
// ===== library types =====

// folder: IO-Link Datatypes/3SU1 IDKey Switch

TYPE "LIOLink_3SU1_IDKeySwitch_typePII"
VERSION : 0.1
   STRUCT
      Status : Byte;
      IDKeyPlugged : Bool;
      AuthLvl_BIT0 : Bool;
      AuthLvl_BIT1 : Bool;
      AuthLvl_BIT2 : Bool;
      SwitchPos_BIT0 : Bool;
      SwitchPos_BIT1 : Bool;
      SwitchPos_BIT2 : Bool;
      Reserved : Bool;
   END_STRUCT;
END_TYPE

// folder: IO-Link ProzessData

TYPE "LIOLink_RF200_typePII"
TITLE = RFID_PII
VERSION : 0.1
   STRUCT
      UID : Array[0..7] of Byte;   // UID capturing / UID Erfassung
   END_STRUCT;
END_TYPE

TYPE "LIOLink_RF200_typePIQ"
TITLE = RFID_PIQ
VERSION : 0.1
   STRUCT
      AntennaOnOff : Byte;   // Antenna switch off with 16#10 (Bit 4 = TRUE) / Antenne ausschalten mit 16#10 (Bit 4 = TRUE)
      reserved : Array[0..6] of Byte;   // Reserved / Reserviert
   END_STRUCT;
END_TYPE

TYPE "LIOLink_3RR24_typePIQ"
TITLE = 3RR24_PIQ
VERSION : 0.1
   STRUCT
      StartOnDelayTime : Bool;   // Start On-Delay time / Starte Anlaufverzögerungszeit
      DQx1 : Bool;   // reserved / Reserviert
      DQx2 : Bool;   // reserved / Reserviert
      Reset : Bool;   // Reset
      DQx4 : Bool;   // reserved / Reserviert
      DQx5 : Bool;   // reserved / Reserviert
      DQx6 : Bool;   // reserved / Reserviert
      DQx7 : Bool;   // reserved / Reserviert
      DQx8 : Bool;   // reserved / Reserviert
      DQx9 : Bool;   // reserved / Reserviert
      DQx10 : Bool;   // reserved / Reserviert
      DQx11 : Bool;   // reserved / Reserviert
      DQx12 : Bool;   // reserved / Reserviert
      DQx13 : Bool;   // reserved / Reserviert
      DQx14 : Bool;   // reserved / Reserviert
      DQx15 : Bool;   // reserved / Reserviert
   END_STRUCT;
END_TYPE

TYPE "LIOLink_3RS1_typePIQ"
TITLE = 3RS14_PIQ
VERSION : 0.1
   STRUCT
      StartOnDelayTime : Bool;   // Start On-Delay time / Starte Anlaufverzögerungszeit
      DQx1 : Bool;   // reserved / Reserviert
      DQx2 : Bool;   // reserved / Reserviert
      Reset : Bool;   // Reset
      DQx4 : Bool;   // reserved / Reserviert
      DQx5 : Bool;   // reserved / Reserviert
      DQx6 : Bool;   // reserved / Reserviert
      DQx7 : Bool;   // reserved / Reserviert
      DQx8 : Bool;   // reserved / Reserviert
      DQx9 : Bool;   // reserved / Reserviert
      DQx10 : Bool;   // reserved / Reserviert
      DQx11 : Bool;   // reserved / Reserviert
      DQx12 : Bool;   // reserved / Reserviert
      DQx13 : Bool;   // reserved / Reserviert
      DQx14 : Bool;   // reserved / Reserviert
      DQx15 : Bool;   // reserved / Reserviert
   END_STRUCT;
END_TYPE

TYPE "LIOLink_3UG48_typePIQ"
TITLE = 3UG48_PIQ
VERSION : 0.1
   STRUCT
      StartTime : Bool;   // Start stabilization or On-Delay time / Starte Stabilisierungs- oder Anlaufverzögerungszeit
      DQx1 : Bool;   // reserved / Reserviert
      DQx2 : Bool;   // reserved / Reserviert
      Reset : Bool;   // Reset
      DQx4 : Bool;   // reserved / Reserviert
      DQx5 : Bool;   // reserved / Reserviert
      DQx6 : Bool;   // reserved / Reserviert
      DQx7 : Bool;   // reserved / Reserviert
      DQx8 : Bool;   // reserved / Reserviert
      DQx9 : Bool;   // reserved / Reserviert
      DQx10 : Bool;   // reserved / Reserviert
      DQx11 : Bool;   // reserved / Reserviert
      DQx12 : Bool;   // reserved / Reserviert
      DQx13 : Bool;   // reserved / Reserviert
      DQx14 : Bool;   // reserved / Reserviert
      DQx15 : Bool;   // reserved / Reserviert
   END_STRUCT;
END_TYPE

TYPE "LIOLink_3RR24_typePII"
TITLE = 3RR24_PII
VERSION : 0.1
// Das Prozessabbild der Eingänge enthält die wichtigsten Statusinformationen der
// Stromüberwachungsrelais 3RR24.
   STRUCT
      Rdy : Bool;   // Ready / Betriebsbereit
      DIx1 : Bool;   // reserved / Reserviert
      GroupError : Bool;   // Group error / Sammelfehler
      GroupWarning : Bool;   // Group warning / Sammelwarnung
      K1 : Bool;   // Status output relay K1 / Status Ausgangrelais K1
      DIx5 : Bool;   // reserved / Reserviert
      DIx6 : Bool;   // reserved / Reserviert
      DIx7 : Bool;   // reserved / Reserviert
      AnalogValueCoding : Byte;   // Analog value coding (only Bit 0..5) / Analogwertcodierung (nur Bit 0..5)
      AnalogValue : Int;   // Analog value / Analogwert
   END_STRUCT;
END_TYPE

TYPE "LIOLink_3UG48_typePII"
TITLE = 3UG48_PII / 3RR24_PII
VERSION : 0.1
// Das Prozessabbild der Eingänge enthält die wichtigsten Statusinformationen der
// Stromüberwachungsrelais 3RR24.
   STRUCT
      Rdy : Bool;   // Ready / Betriebsbereit
      DIx1 : Bool;   // reserved / Reserviert
      GroupError : Bool;   // Group error / Sammelfehler
      GroupWarning : Bool;   // General or group warning / Sammelwarnung
      K1 : Bool;   // Status output relay K1 / Status Ausgangrelais K1
      DIx5 : Bool;   // reserved / Reserviert
      DIx6 : Bool;   // reserved / Reserviert
      DIx7 : Bool;   // reserved / Reserviert
      AnalogValueCoding : Byte;   // Analog value coding (only Bit 0..5) / Analogwertcodierung (nur Bit 0..5)
      AnalogValue : Int;   // Analog value / Analogwert
   END_STRUCT;
END_TYPE

TYPE "LIOLink_3RA_typePII"
TITLE = 3RAxy_PII
VERSION : 0.1
// Data Type of the process input image contains the important status information of all compact starters. / Datentyp für das Prozessabbild der Eingänge enthält die wichtigen Statusinformationen aller Kompaktabzweige.
   STRUCT
      St1Rdy : Bool;   // Starter 1 ready (automatic) / Starter 1 Bereit (Automatik)
      St1MotorOn : Bool;   // Starter 1 Motor on / Starter 1 Motor ein
      St1Fault : Bool;   // Starter 1 group fault / Starter 1 Sammelfehler
      St1Warn : Bool;   // Starter 1 group warning / Starter 1 Sammelwarnung
      St2Rdy : Bool;   // Starter 2 ready (automatic) / Starter 2 Bereit (Automatik)
      St2MotorOn : Bool;   // Starter 2 Motor on / Starter 2 Motor ein
      St2Fault : Bool;   // Starter 2 group fault / Starter 2 Sammelfehler
      St2Warn : Bool;   // Starter 2 group warning / Starter 2 Sammelwarnung
      St3Rdy : Bool;   // Starter 3 ready (automatic) / Starter 3 Bereit (Automatik)
      St3MotorOn : Bool;   // Starter 3 Motor on / Starter 3 Motor ein
      St3Fault : Bool;   // Starter 3 group fault / Starter 3 Sammelfehler
      St3Warn : Bool;   // Starter 3 group warning / Starter 3 Sammelwarnung
      St4Rdy : Bool;   // Starter 4 ready (automatic) / Starter 4 Bereit (Automatik)
      St4MotorOn : Bool;   // Starter 4 Motor on / Starter 4 Motor ein
      St4Fault : Bool;   // Starter 4 group fault / Starter 4 Sammelfehler
      St4Warn : Bool;   // Starter 4 group warning / Starter 4 Sammelwarnung
   END_STRUCT;
END_TYPE

TYPE "LIOLink_3RA_typePIQ"
TITLE = 3RAxy_PIQ
VERSION : 0.1
// The process output image contains the control commands for all compact starters. / Datentyp für das Prozessabbild der Ausgänge enthält die Steuerbefehle für alle Kompaktabzweige.
   STRUCT
      St1Dir1 : Bool;   // Starter 1 Motor direction of rotation 1 / Starter 1 Motor Drehrichtung 1
      St1Dir2 : Bool;   // Starter 1 Motor direction of rotation 2 / Starter 1 Motor Drehrichtung 2
      St1Res : Bool;   // Starter 1 Reserved / Starter 1 reserviert
      St1TripReset : Bool;   // Starter 1 Trip reset / Starter 1 Trip-Reset
      St2Dir1 : Bool;   // Starter 2 Motor direction of rotation 1 / Starter 2 Motor Drehrichtung 1
      St2Dir2 : Bool;   // Starter 2 Motor direction of rotation 2 / Starter 2 Motor Drehrichtung 2
      St2Res : Bool;   // Starter 2 Reserved / Starter 2 reserviert
      St2TripReset : Bool;   // Starter 2 Trip reset / Starter 2 Trip-Reset
      St3Dir1 : Bool;   // Starter 3 Motor direction of rotation 1 / Starter 3 Motor Drehrichtung 1
      St3Dir2 : Bool;   // Starter 3 Motor direction of rotation 2 / Starter 3 Motor Drehrichtung 2
      St3Res : Bool;   // Starter 3 Reserved / Starter 3 reserviert
      St3TripReset : Bool;   // Starter 3 Trip reset / Starter 3 Trip-Reset
      St4Dir1 : Bool;   // Starter 4 Motor direction of rotation 1 / Starter 4 Motor Drehrichtung 1
      St4Dir2 : Bool;   // Starter 4 Motor direction of rotation 2 / Starter 4 Motor Drehrichtung 2
      St4Res : Bool;   // Starter 4 Reserved / Starter 4 reserviert
      St4TripReset : Bool;   // Starter 4 Trip reset / Starter 4 Trip-Reset
   END_STRUCT;
END_TYPE

TYPE "LIOLink_3RB24_typePII"
TITLE = 3RB24_PII
VERSION : 0.1
// Data Type of the process input image contains the most important status information of the solid-state overload relay for IO‑Link.
// Datentyp für das Prozessabbild der Eingänge enthält die wichtigsten Statusinformationen des
// elektronischen Überlastrelais für IO-Link.
   STRUCT
      Rdy : Bool;   // Ready (automatic) / Bereit (Automatik)
      MotorOn : Bool;   // Motor on / Motor ein
      GroupFault : Bool;   // Group fault / Sammelfehler
      GroupWarning : Bool;   // Group warning / Sammelwarnung
      DIx4 : Bool;   // reserved / reserviert
      DIx5 : Bool;   // reserved / reserviert
      DIx6 : Bool;   // reserved / reserviert
      DIx7 : Bool;   // reserved / reserviert
      CurrentRatio : Byte;   // Bit 0..5: Motor current ratio (%), Bit 6: Manual mode / Bit 0..5: Motorstromverhältnis, Bit 6: Handbetrieb
   END_STRUCT;
END_TYPE

TYPE "LIOLink_3RB24_typePIQ"
TITLE = 3RB24_PIQ
VERSION : 0.1
// The process output image contains the control commands for the solid-state overload relay for IO‑Link.
// Datentyp für das Prozessabbild der Ausgänge enthält die Steuerbefehle für das elektronische
// Überlastrelais für IO-Link
   STRUCT
      Direction1 : Bool;   // Motor direction of rotation 1 / Motor Drehrichtung 1
      Direction2 : Bool;   // Motor direction of rotation 2 / Motor Drehrichtung 2
      DQx2 : Bool;   // Reserved / reserviert
      TripReset : Bool;   // Trip reset / Trip-Reset
      DQx4 : Bool;   // Reserved / reserviert
      DQx5 : Bool;   // Reserved / reserviert
      DQx6 : Bool;   // Reserved / reserviert
      DQx7 : Bool;   // Reserved / reserviert
      DQx8 : Bool;   // Reserved / reserviert
      DQx9 : Bool;   // Reserved / reserviert
      DQx10 : Bool;   // Reserved / reserviert
      DQx11 : Bool;   // Reserved / reserviert
      DQx12 : Bool;   // Reserved / reserviert
      DQx13 : Bool;   // Reserved / reserviert
      DQx14 : Bool;   // Reserved / reserviert
      DQx15 : Bool;   // Reserved / reserviert
   END_STRUCT;
END_TYPE

TYPE "LIOLink_3RS1_typePII"
TITLE = 3RS14_PII
VERSION : 0.1
   STRUCT
      Rdy : Bool;   // Ready / Betriebsbereit
      DIx1 : Bool;   // reserved / Reserviert
      GroupError : Bool;   // Group error / Sammelfehler
      GroupWarning : Bool;   // General or group warning / Sammelwarnung
      K1 : Bool;   // Status output relay K1 / Status Ausgangrelais K1
      K2 : Bool;   // Status output relay K2 / Status Ausgangrelais K2
      K3 : Bool;   // Status output relay K3 / Status Ausgangrelais K3
      DIx7 : Bool;   // reserved / Reserviert
      AnalogValueCoding : Byte;   // Analog value coding (only Bit 0..4) / Analogwertcodierung (nur Bit 0..4)
      AnalogValue : Int;   // Analog value / Analogwert
   END_STRUCT;
END_TYPE

// folder: LIOLink

TYPE "LIOLink_typeDiagnostics"
   STRUCT
      status : Word;   // Status of the Block or error identification when error occurred
      subfunctionStatus : DWord;   // Status or return value of called FB's, FCs and system blocks
      stateNumber : DInt;   // State in the state machine of the block where the error occurred
   END_STRUCT;
END_TYPE

// folder: LIOLink/Common

TYPE "LIOLink_typePortEventQualifier"
TITLE = LIOLink_typePortEventQualifier
// EventQualifier: Instance, Source, Type, Mode
   STRUCT
      instance : Byte;   // 0: Unknown / 1-3: Reserved / 4: Application / 5-7: Reserved
      source : Bool;   // (default) FALSE: Device (remote) / TRUE: Master/Port
      "type" : Byte;   // 0: Reserved / 1: Notification / 2: Warning / 3: Error
      mode : Byte;   // 0: Reserved / 1: Event single shot / 2: Event disappears / 3: Event appears
   END_STRUCT;
END_TYPE

TYPE "LIOLink_typePortEventCodes"
TITLE = LIOLink_PortEventCodes
// UDT for Event Information: eventCode, eventQualifier
   STRUCT
      eventCode : Word;   // IO-Link EventCode
      eventQualifier : "LIOLink_typePortEventQualifier";   // IO-Link EventQualifier
   END_STRUCT;
END_TYPE

TYPE "LIOLink_typePortEvents"
TITLE = LIOLink_PortEvents
// Events of a port
   STRUCT
      event : Array[0..4] of "LIOLink_typePortEventCodes";   // Events of a port
   END_STRUCT;
END_TYPE

TYPE "LIOLink_typeEvents"
TITLE = LIOLink_Events
// Events of each port of a IO-Link-Master
   STRUCT
      port : Array[1..8] of "LIOLink_typePortEvents";   // Ports of IO-Link-Master
   END_STRUCT;
END_TYPE

// folder: LIOLink/Common/Device-specific data types/SIMATIC RF200

TYPE "LIOLink_RF200_typeParameters"
TITLE = LIOLink_RF200_typeParameters
// Contains all parameters of a RF200
   STRUCT
      eventMessage : Byte;   // 16#02: Event indication enabled (default), 16#04: No Message
      operatingMode : Byte;   // 16#04: Scan UID (default), 16#08 Scan user data
      readyDelay : Byte;   // 16#02 Turn off (default), 16#04: Turn on additional backup mechanism for
      dataHoldingTime : Byte;   // Minimum time during which the process input data is not changed by the device
      rfParameters : Byte;   // Setting the RF parameters, 16#02 ISO default, 16#04: special settings
      modulation : Byte;   // Setting for the modulation strength 16#00 (0%) ... 16#64 (100%) - default 16#16 (22%)
      subcarrier : Byte;   // Subcarrier, 16#02: Single (default), 16#04: double
      dataTransfer : Byte;   // Data transmission speed, 16#02: low, 16#04: high (default)
   END_STRUCT;
END_TYPE

TYPE "LIOLink_RF200_typeEventHistory"
TITLE = LIOLink_RF200_typeEventHistory
VERSION : 0.1
// Contains last 5 events of a RF200
   STRUCT
      lastEvent : DWord;   // Last event
      secondLastEvent : DWord;   // Second last event
      thirdLastEvent : DWord;   // Third last event
      fourthLastEvent : DWord;   // Fourth last event
      fifthLastEvent : DWord;   // Fifth last event
   END_STRUCT;
END_TYPE

TYPE "LIOLink_RF200_typeReaderStatus"
TITLE = LIOLink_RF200_typeReaderStatus
VERSION : 0.1
// Contrains all information about the status of the reader
   STRUCT
      timeSinceStartup : DWord;   // Operating time in seconds
      tagsInTheField : Byte;   // current number of transponders in the field
      antennaStatus : Byte;   // antenna turned on/off
      tagChanges : DWord;   // number of transponder changes
      lineDriverRev : Byte;   // version of the IO-Link line driver
      errorCounterPassive : Byte;   // Air interface: Counter for errors in idle state
      abortCounter : Byte;   // Air interface: Communication aborted
      codeErrorCounter : Byte;   // Air interface: Communication disruption
      signatureErrorCounter : Byte;   // Air interface: Protocol error, signature error counter, is reset when read out
      crcErrorCounter : Byte;   // Air interface: Communication disruption
      currentCommandStatus : Byte;   // Command status of the last command, is reset when read out
      errorCount : Byte;   // HOST interface: Communication disruption
   END_STRUCT;
END_TYPE

TYPE "LIOLink_RF200_typeUIDHistory"
TITLE = LIOLink_RF200_typeUIDHistory
VERSION : 0.1
// Contains UID history
   STRUCT
      lastUID1 : DWord;   // Last UID
      lastUID2 : DWord;   // Last UID
      secondLastUID1 : DWord;   // Second last UID
      secondLastUID2 : DWord;   // Second last UID
      thirdLastUID1 : DWord;   // Third last UID
      thirdLastUID2 : DWord;   // Third last UID
      fourthLastUID1 : DWord;   // Fourth last UID
      fourthLastUID2 : DWord;   // Fourth last UID
      fifthLastUID1 : DWord;   // Fifth last UID
      fifthLastUID2 : DWord;   // Fifth last UID
   END_STRUCT;
END_TYPE

TYPE "LIOLink_RF200_typeTagStatus"
TITLE = LIOLink_RF200_typeTagStatus
VERSION : 0.1
// Contains all the information about the status of the tag
   STRUCT
      uid : Array[0..7] of Byte;   // Unique identifier of the transponder
      tagName : Byte;   // Transponder Name
      chipVersion : Byte;   // Version of the Chip
      memSize : Word;   // Memory size in Bytes
      lockStatus : Byte;   // Disable blocks on the chip
      memBlockSize : Byte;   // Size of memory blocks of the chip
      numBlocks : Byte;   // Number of memory blocks of the chip
   END_STRUCT;
END_TYPE

TYPE "LIOLink_RF200_typeAll"
TITLE = LIOLink_RF200_typeAll
VERSION : 0.1
// Contains all information about RF200
   STRUCT
      directParameterPage : "LIOLink_typeParameterPage0";   // ID0: Parameter page 0
      systemCommand : Byte;   // ID2: System command
      deviceAccessLocks : Word;   // ID12: Device access locks
      vendorName : String[12];   // ID16: Vendor name
      vendorText : String[12];   // ID17: Vendor text
      productName : String[24];   // ID18: Product name
      productID : String[16];   // ID19: Product ID
      productText : String[64];   // ID20: Product Text
      serialNumber : String[12];   // ID21: Serial Number
      hwRevision : String[12];   // ID22: Hardware revision
      fwRevision : String[12];   // ID23: Firmware revision
      appSpecificName : String[32];   // ID24: Application specific name
      errorCount : Word;   // ID32: Number of errors that have occured (not warnings)
      deviceStatus : Byte;   // ID36: Device status
      deviceStatusDetailed : Byte;   // ID37: Detailed device status
      processImageIn : Array[0..7] of Byte;   // ID40: Read out last process image of the inputs
      processImageOut : Array[0..7] of Byte;   // ID41: Read out last process image of the outputs
      parameters : "LIOLink_RF200_typeParameters";   // ID64: Read/Write Reader Parameters
      eventHistory : "LIOLink_RF200_typeEventHistory";   // ID74: Number of events
      readerStatus : "LIOLink_RF200_typeReaderStatus";   // ID90: Reader status
      tagStatus : "LIOLink_RF200_typeTagStatus";   // ID91: Tag status
      uidHistory : "LIOLink_RF200_typeUIDHistory";   // ID92: History of UID
   END_STRUCT;
END_TYPE

// folder: LIOLink/Common/Device-specific data types/SIRIUS/3RA

TYPE "LIOLink_3RA_typeDiagStarterShort"
TITLE = LIOLink_3RA_typeDiagStarterShort
// Contains diagnose of starter of type "short"
   STRUCT
      starterItemNumber : Byte;   // Starter Item number (1 to 4)
      starterAvailable : Byte;   // Starter Available: 16#00 not available; 16#02: available
      reserved1 : Array[2..5] of Byte;   // Reserved
      contactBlockDefective : Bool;   // Contact block defective
      contactSupplyVoltageMissing : Bool;   // Contact block supply voltage missing
      reserved2 : Bool;   // Reserved
      trippMotorOverload : Bool;   // Motor overload tripping
      trippCircuitBreaker : Bool;   // Circuit breaker tripped
      switchOffendPosRight : Bool;   // Switch off - end position right
      switchOffendPosLeft : Bool;   // Switch off - end position left
      processImageError : Bool;   // Process image error
      manualOperationLocal : Bool;   // Manual operation local
      manualOperationConAborted : Bool;   // Manual operation connection aborted
      ContactCoolingTimeActive : Bool;   // Contact block cooling time active
      remainingLifeTime0 : Bool;   // Remaining life time (RLT 0%)
      reserved3 : Bool;   // Reserved
      reserved4 : Bool;   // Reserved
      reserved5 : Bool;   // Reserved
      reserved6 : Bool;   // Reserved
   END_STRUCT;
END_TYPE

TYPE "LIOLink_3RA_typeDiagStarterLong"
TITLE = LIOLink_3RA_typeDiagStarterLong
// Contains diagnose of starter of type "long"
   STRUCT
      reserved1 : Byte;   // Reserved
      starterItemNumber : Byte;   // Starter Item number (1 to 4)
      starterAvailable : Byte;   // Starter Available: 16#00 not available; 16#02: available
      reserved2 : Array[3..6] of Byte;   // Reserved
      contactBlockDefective : Bool;   // Contact block defective
      contactSupplyVoltageMissing : Bool;   // Contact block supply voltage missing
      reserved3 : Bool;   // Reserved
      trippMotorOverload : Bool;   // Motor overload tripping
      trippCircuitBreaker : Bool;   // Circuit breaker tripped
      switchOffendPosRight : Bool;   // Switch off - end position right
      switchOffendPosLeft : Bool;   // Switch off - end position left
      processImageError : Bool;   // Process image error
      manualOperationLocal : Bool;   // Manual operation local
      manualOperationConAborted : Bool;   // Manual operation connection aborted
      ContactCoolingTimeActive : Bool;   // Contact block cooling time active
      remainingLifeTime0 : Bool;   // Remaining life time (RLT 0%)
      reserved4 : Bool;   // Reserved
      reserved5 : Bool;   // Reserved
      reserved6 : Bool;   // Reserved
      reserved7 : Bool;   // Reserved
      reserved8 : Byte;   // Reserved
   END_STRUCT;
END_TYPE

TYPE "LIOLink_3RA_typeConfigStarterShort"
TITLE = LIOLink_3RA_typeConfigStarterShort
// Contains configurations for starter with type "short"
   STRUCT
      starterItemNumber : Byte;   // Starter (item number)
      reserved1 : Byte := 16#60;   // Fixed Value
      starterDiag : Byte;   // Starter Diag: 16#00: not available; 16#02: available but defect; 16#03: available and OK
      starterType : Byte;   // Type of starter
      starterVersion1 : Byte;   // Starter Version part 1
      starterVersion2 : Byte;   // Starter Version part 2
   END_STRUCT;
END_TYPE

TYPE "LIOLink_3RA_typeConfigStarterLong"
TITLE = LIOLink_3RA_typeConfigStarterLong
// Contains configurations for starter with type "long"
   STRUCT
      reserved : Byte := 16#07;   // Fixed Value
      starterItemNumber : Byte;   // Starter (item number)
      reserved1 : Byte := 16#60;   // Fixed Value
      starterDiag : Byte;   // Starter Diag: 16#00: not available; 16#02: available but defect; 16#03: available and OK
      starterType : Byte;   // Type of starter
      starterVersion1 : Byte;   // Starter Version part 1
      starterVersion2 : Byte;   // Starter Version part 2
      reserved2 : Byte := 16#07;   // Fixed Value
   END_STRUCT;
END_TYPE

TYPE "LIOLink_3RA_typeDiag"
TITLE = LIOLink_3RA_typeDiag
VERSION : 0.1
// Data set (index) 90 - group diagnostics: Starter group
   STRUCT
      reserved : Array[0..3] of Byte;   // Reserved - Dataset Index 90 - Length 53 / read length 52
      numberOfStarters : Byte;   // Number of starters (compact starters and operator panel)
      configurationCompare : Byte;   // Preset <> actual configuration 16#00: equal 16#01: different
      reserved1 : Word;   // Reserved
      starter1 : "LIOLink_3RA_typeDiagStarterLong";   // Starter 1 - module and specific diagnostics
      starter2 : "LIOLink_3RA_typeDiagStarterShort";   // Starter 2 - module and specific diagnostics
      starter3 : "LIOLink_3RA_typeDiagStarterLong";   // Starter 3 - module and specific diagnostics
      starter4 : "LIOLink_3RA_typeDiagStarterShort";   // Starter 4 - module and specific diagnostics
      reserved3 : Byte;   // Reserved
      operatorItemNumber : Byte;   // Operator panel (item number)
      operatorAvailable : Byte;   // Operator panel available: 16#00 not available; 16#02: available
      reserved4 : Byte;   // Reserved
      reserved5 : Array[48..51] of Byte;   // Reserved
   END_STRUCT;
END_TYPE

TYPE "LIOLink_3RA_typeConfig"
TITLE = LIOLink_3RA_typeConfig / IO-Link Parameter mit dem Baustein "FB IO_CALL" auslesen!
VERSION : 0.1
// Contains all the possible configurations of 3RA
   STRUCT
      reserved : Array[0..7] of Byte;   // Reserved
      starter1 : "LIOLink_3RA_typeConfigStarterLong";   // Config Data of Starter 1
      starter2 : "LIOLink_3RA_typeConfigStarterShort";   // Config Data of Starter 2
      starter3 : "LIOLink_3RA_typeConfigStarterLong";   // Config Data of Starter 3
      starter4 : "LIOLink_3RA_typeConfigStarterShort";   // Config Data of Starter 4
      reserved1 : Byte := 16#07;   // Reserved
      operatorItemNumber : Byte;   // Operator panel (item number)
      reserved2 : Byte := 16#60;   // Reserved
      operatorAvailable : Byte;   // Operator panel available: 16#00 not available; 16#02: available
      reserved3 : Byte := 16#D2;   // Reserved
      reserved4 : Byte;   // Reserved
   END_STRUCT;
   // reserved[0] := 16#0021;
   // reserved[1] := 16#0000;
   // reserved[2] := 16#0000;
   // reserved[3] := 16#0000;
   // reserved[4] := 16#0005;
END_TYPE

TYPE "LIOLink_3RA_typeAll"
TITLE = LIOLink_3RA_typeAll
VERSION : 0.1
// Contains all the information about 3RA
   STRUCT
      parameterPage0 : "LIOLink_typeParameterPage0";   // ID0: Parameter page 0
      parameterPage1 : "LIOLink_3RA_typeParameterPage1";   // ID1: Parameter page 1
      vendorName : String[10];   // ID16: Vendor name
      vendorText : String[58];   // ID17: Vendor text
      productName : String[30];   // ID18: Product name
      productID : String[8];   // ID19: Product ID
      productText : String[2];   // ID20: Product text
      serialNumber : String[8];   // ID21: Serial number
      hwRevision : String[4];   // ID22: Hardware revision
      fwRevision : String[4];   // ID23: Firmware revision
      appSpecificName : String[32];   // ID24: Application specific name
      diagnostics : "LIOLink_3RA_typeDiag";   // ID90: Group diagnostics
      actualConfig : "LIOLink_3RA_typeConfig";   // ID105: Actual configuration
      targetConfig : "LIOLink_3RA_typeConfig";   // ID130: Target configuration
   END_STRUCT;
   // actualConfig.reserved[0] := 16#0021;
   // actualConfig.reserved[1] := 16#0000;
   // actualConfig.reserved[2] := 16#0000;
   // actualConfig.reserved[3] := 16#0000;
   // actualConfig.reserved[4] := 16#0005;
   // targetConfig.reserved[0] := 16#0021;
   // targetConfig.reserved[1] := 16#0000;
   // targetConfig.reserved[2] := 16#0000;
   // targetConfig.reserved[3] := 16#0000;
   // targetConfig.reserved[4] := 16#0005;
END_TYPE

TYPE "LIOLink_3RA_typeParameterPage1"
TITLE = LIOLink_3RA_typeParameterPage1 / IO-Link Parameter mit dem Baustein "FB IO_CALL" auslesen!
AUTHOR : SIE_RS
FAMILY : 3RA
NAME : IO-Link
VERSION : 1.0
// Contains Parameter Page 1 of 3RA
   STRUCT
      productFamiliy : Byte;   // Produktfamily SIRIUS (0x60) - A-9 Dataset Index 1 Page 75
      starter1Compare : Bool;   // Starter 1 - 0: Target/actual comparison: Yes, 1: Target/actual comparison: No,
      starter1Available : Bool;   // Starter 1 - 0: Starter available: No, 1: Starter available: Yes,
      starter2Compare : Bool;   // Starter 2 - 0: Target/actual comparison: Yes, 1: Target/actual comparison: No,
      starter2Available : Bool;   // Starter 2 - 0: Starter available: No, 1: Starter available: Yes,
      starter3Compare : Bool;   // Starter 3 - 0: Target/actual comparison: Yes, 1: Target/actual comparison: No,
      starter3Available : Bool;   // Starter 3 - 0: Starter available: No, 1: Starter available: Yes,
      starter4Compare : Bool;   // Starter 4 - 0: Target/actual comparison: Yes, 1: Target/actual comparison: No,
      starter4Available : Bool;   // Starter 4 - 0: Starter available: No, 1: Starter available: Yes,
      operatorPanelCompare : Bool;   // Operator panel - 0:Target/actual comparison: Yes, 1:Target/actual comparison:No
      operatorPanelAvailable : Bool;   // Operator panel - 0: Starter available: No, 1: Starter available: Yes,
      reserved1 : Bool;   // Reserved
      reserved2 : Bool;   // Reserved
      profileVersion1 : Bool;   // Profile version
      profileVersion2 : Bool;   // Profile version
      profileVersion3 : Bool;   // Profile version
      profileVersion4 : Bool;   // Profile version
      starter1Type : Byte;   // Starter 1 - Type of starter
      starter1Version : Byte;   // Starter 1 - Starter version
      starter2Type : Byte;   // Starter 2 - Type of starter
      starter2Version : Byte;   // Starter 2 - Starter version
      starter3Type : Byte;   // Starter 3 - Type of starter
      starter3Version : Byte;   // Starter 3 - Starter version
      starter4Type : Byte;   // Starter 4 - Type of starter
      starter4Version : Byte;   // Starter 4 - Starter version
      operatorPanel : Byte;   // 210: Operator panel
      reserved3 : Byte;   // Reserved
      reserved4 : Byte;   // Reserved
      reserved5 : Byte;   // Reserved
      reserved6 : Byte;   // Reserved
   END_STRUCT;
END_TYPE

// folder: LIOLink/Common/Device-specific data types/SIRIUS/3RB24

TYPE "LIOLink_3RB24_typeMeasure"
TITLE = LIOLink_3RB24_typeMeasure
VERSION : 0.1
// Data set (index) 94 (measured values) - solid-state overload relay for IO‑Link
   STRUCT
      phaseCurrentL1Rel : Byte;   // Phase current I (L1 rms in 3,125% steps) - A-4 Dataset Index 94 Page 112
      phaseCurrentL2Rel : Byte;   // Phase current I (L2 rms in 3,125 % steps)
      phaseCurrentL3Rel : Byte;   // Phase current I (L3 rms in 3,125 % steps)
      reserved : Byte;   // Reserved
      reserved1 : Array[4..27] of Byte;   // Reserved
      phaseCurrentL1Abs : DWord;   // Phase current I (L1 rms in 0,01-A steps)
      phaseCurrentL2Abs : DWord;   // Phase current I (L2 rms in 0,01-A steps)
      phaseCurrentL3Abs : DWord;   // Phase current I (L3 rms in 0,01-A steps)
   END_STRUCT;
END_TYPE

TYPE "LIOLink_3RB24_typeTechFunctions"
TITLE = TechnologyFunctions_3RB24
VERSION : 0.1
// Data set (index) 131 (technology functions) - solid-state overload relay for IO‑Link
   STRUCT
      reserved : Array[0..7] of Byte;   // Reserved
      groundFaultDetection : Byte;   // Ground fault detection - 16#00: Disable; 16#20: Enable - Bit 5 in Byte
      reserved8 : Word;   // Reserved
      coldStart : Byte;   // Cold Start - 16#00: Disable; 16#08: Enable - Bit 3 in Byte
      ratedOpCurrent : DWord;   // Rated operational current (in 0.01 A steps)
      reserved16 : Word;   // Reserved
      responseToOverloadMotor : Byte;   // Response to overload - thermal motor model - 16#00: Tripping without restart (MAN); 16#01: Tripping with restart (AUTO)
      tripClass : Byte;   // Trip class - 16#03: CLASS 5; 16#00: CLASS 10; 16#01: CLASS 20; 16#02: CLASS 30
      reserved17 : DWord;   // Reserved
      responseToOverloadThermistor : Bool;   // Response to overload - Thermistor - false: Tripping without restart (MAN); true: Tripping with restart (AUTO)
      reserved18 : Bool;   // Reserved
      reserved19 : Bool;   // Reserved
      reserved20 : Bool;   // Reserved
      reserved21 : Bool;   // Reserved
      reserved22 : Bool;   // Reserved
      reserved23 : Bool;   // Reserved
      monitorThermistor : Bool;   // Thermistor - monitoring - false: No; true: Yes
   END_STRUCT;
END_TYPE

TYPE "LIOLink_3RB24_typePresetConfig"
TITLE = TargetConfiguration_3RB24
VERSION : 0.1
// Data set (index) 130 (target configuration) - operator panel
   STRUCT
      reserverd : Array[0..17] of Byte;   // Reserved
      reserved1 : Bool;   // Reserved
      reserved2 : Bool;   // Reserved
      reserved3 : Bool;   // Reserved
      reserved4 : Bool;   // Reserved
      reserved5 : Bool;   // Reserved
      reserved6 : Bool;   // Reserved
      operationAtTarget : Bool;   // Operation at Preset <> Actual Configuration
      operationPanelAvailable : Bool;   // Operator panel available
      reserved7 : Byte;   // Reserved
      reserved8 : Byte;   // Reserved
      reserved9 : Byte;   // Reserved
   END_STRUCT;
END_TYPE

TYPE "LIOLink_3RB24_typeDiag"
TITLE = LIOLink_3RB24_typeDiag
VERSION : 0.1
// Data set (index) 94 (measured values) - solid-state overload relay for IO‑Link
   STRUCT
      ready : Bool;   // Ready
      directionClockwise : Bool;   // Motor direction of rotation 1 (clockwise)
      directionCounterClockwise : Bool;   // Motor direction of rotation 2 (counter-clockwise)
      reserved : Bool;   // Reserved
      switchingElementDefect : Bool;   // Switching element defective
      reserved1 : Bool;   // Reserved
      groupError : Bool;   // GroupError
      generalWarning : Bool;   // General warning
      reserved2 : Byte;   // Reserved
      thermistorOverload : Bool;   // Thermistor overload
      thermistorWireBreak : Bool;   // Thermistor wire break
      thermistorShortCircuit : Bool;   // Thermistor short-circuit
      thermistorMotorOverload : Bool;   // Thermal motor model overload
      overloadTripping : Bool;   // Overload tripping
      reserved3 : Bool;   // Reserved
      reserved4 : Bool;   // Reserved
      reserved5 : Bool;   // Reserved
      reserved6 : Byte;   // Reserved
      reserved7 : Bool;   // Reserved
      reserved8 : Bool;   // Reserved
      reserved9 : Bool;   // Reserved
      reserved10 : Bool;   // Reserved
      reserved11 : Bool;   // Reserved
      resCurrenctDetected : Bool;   // Residual current detected
      resCurrentTripping : Bool;   // Residual current tripping
      reserved12 : Bool;   // Reserved
      reserved13 : Byte;   // Reserved
      groudFaultDetected : Bool;   // Ground fault detected
      GroundFaultTripping : Bool;   // Ground fault tripping
      reserved14 : Bool;   // Reserved
      reserved15 : Bool;   // Reserved
      reserved16 : Bool;   // Reserved
      reserved17 : Bool;   // Reserved
      reserved18 : Bool;   // Reserved
      supplyVoltageLow : Bool;   // Electronics supply voltage too low
      reserved19 : Bool;   // Reserved
      reserved20 : Bool;   // Reserved
      autoMode1 : Bool;   // Automatic mode
      autoMode2 : Bool;   // Automatic mode
      manualModeOP1 : Bool;   // Manual mode (operator panel)
      manualModeOP2 : Bool;   // Manual mode (operator panel)
      manualModeConAbort : Bool;   // Manual mode connection abort (operator panel)
      processImageError : Bool;   // Process image error
      reserved21 : Byte;   // Reserved
      selfTestActive1 : Bool;   // Self-test active
      selfTestActive2 : Bool;   // Self-test active
      selfTestError : Bool;   // Self-test error
      reserved22 : Bool;   // Reserved
      reserved23 : Bool;   // Reserved
      reserved24 : Bool;   // Reserved
      reserved25 : Bool;   // Reserved
      reserved26 : Bool;   // Reserved
      reserved27 : Word;   // Reserved
      reserved28 : Bool;   // Reserved
      reserved29 : Bool;   // Reserved
      impermissibleSetting : Bool;   // Impermissible Ie/CLASS setting
      presetActualCompare : Bool;   // Preset <> actual configuration
      thermistorProtectionDeactivated : Bool;   // Thermistor protection deactivated
      reserved30 : Bool;   // Reserved
      reserved31 : Bool;   // Reserved
      reserved32 : Bool;   // Reserved
      reserved33 : Byte;   // Reserved
      coldStartActive : Bool;   // Cold start active
      coldStartTripping : Bool;   // Cold start tripping
      reserved34 : Bool;   // Reserved
      reserved35 : Bool;   // Reserved
      reserved36 : Bool;   // Reserved
      reserved37 : Bool;   // Reserved
      reserved38 : Bool;   // Reserved
      reserved39 : Bool;   // Reserved
      reserved40 : Byte;   // Reserved
      reserved41 : Array[16..23] of Byte;   // Reserved
      reserved42 : Bool;   // Reserved
      reserved43 : Bool;   // Reserved
      reserved44 : Bool;   // Reserved
      motorHeatingExceeded : Bool;   // Prewarning limit: Motor heating exceeded
      reserved45 : Bool;   // Reserved
      reserved46 : Bool;   // Reserved
      reserved47 : Bool;   // Reserved
      reserved48 : Bool;   // Reserved
      reserved49 : Byte;   // Reserved - Extension to get even field
   END_STRUCT;
END_TYPE

TYPE "LIOLink_3RB24_typeAll"
TITLE = LIOLink_3RB24_typeAll
VERSION : 0.1
// Contains all the information about 3RB24
   STRUCT
      parameterPage0 : "LIOLink_typeParameterPage0";   // ID0: Parameter page 0
      vendorName : String[10];   // ID16: Vendor name
      vendorText : String[64];   // ID17: Vendor text
      productName : String[30];   // ID18: Product name
      productID : String[12];   // ID19: Product ID
      productText : String[2];   // ID20: Product text
      serialNumber : String[8];   // ID21: Serial number
      hwRevision : String[4];   // ID22: Hardware revision
      fwRevision : String[4];   // ID23: Firmware revision
      appSpecificName : String[32];   // ID24: Application specific name
      processInput : Word;   // ID40: Process data input
      processOutput : Byte;   // ID41: Process data output
      diagnostics : "LIOLink_3RB24_typeDiag";   // ID92: Diagnostics
      measuredValues : "LIOLink_3RB24_typeMeasure";   // ID94: Measurement values
      presetConfig : "LIOLink_3RB24_typePresetConfig";   // ID130: Preset configuration
      techFunctions : "LIOLink_3RB24_typeTechFunctions";   // ID131: Technology functions
   END_STRUCT;
END_TYPE

// folder: LIOLink/Common/Device-specific data types/SIRIUS/3RR24

TYPE "LIOLink_3RR24_typeDiag"
TITLE = LIOLink_3RR24_typeDiag
VERSION : 0.1
// Data set (index) 92 - diagnostics
   STRUCT
      reserved : Array[0..15] of Byte;   // Reserved
      ready : Bool;   // Ready
      groupError : Bool;   // Group error
      groupWarning : Bool;   // Group warning
      reserved1 : Bool;   // Reserved
      reserved2 : Bool;   // Reserved
      parameterAssign : Bool;   // Parameter assignment active
      parameterInvalid : Bool;   // Invalid parameter
      internalError : Bool;   // Self-test error/internal error
      reserved3 : Byte;   // Reserved
      errorNumber : Word;   // Parameter error number
      reserved4 : Array[20..25] of Byte;   // Reserved
      delayTimeRunning : Bool;   // ON-delay time running
      delayLevelUp : Bool;   // Tripping delay time running (threshold for overshoot)
      delayLevelDown : Bool;   // Tripping delay time running (threshold for undershoot)
      delayAsymmetry : Bool;   // Tripping delay time running (threshold for current asymmetry)
      delayReclosing : Bool;   // Reclosing delay time is running
      reserved5 : Bool;   // Reserved
      reserved6 : Bool;   // Reserved
      reserved7 : Bool;   // Reserved
      levelUp : Bool;   // Threshold for overshoot exceeded
      levelDown : Bool;   // Threshold for underhsoot violated
      currentAsymmetry : Bool;   // Threshold for current asymmetry exceeded
      warningLevelUp : Bool;   // Warning threshold for overshoot exceeded
      warningLevelDown : Bool;   // Warning threshold for undershoot violated
      warningCurrentAsymmetry : Bool;   // Warning threshold for current asymmetry exceedd
      reserved8 : Bool;   // Reserved
      reserved9 : Bool;   // Reserved
      reserved10 : Bool;   // Reserved
      phaseFailureL1 : Bool;   // Phase failure L1
      phaseFailureL2 : Bool;   // Phase failure L2
      phaseFailureL3 : Bool;   // Phase failure L3
      overcurrentL1 : Bool;   // Overcurrent n x Imax L1
      overcurrentL2 : Bool;   // Overcurrent n x Imax L2
      overcurrentL3 : Bool;   // Overcurrent n x Imax L3
      reserved11 : Bool;   // Reserved
      faultCurrentExceeded : Bool;   // Threshold for fault current exceeded
      phaseSeqL1L2L3 : Bool;   // Phase sequence L1-L2-L3
      phaseSeqL3L2L1 : Bool;   // Phase sequence L3-L2-L1
      phaseSeqError : Bool;   // Phase sequence error
      reserved12 : Bool;   // Reserved
      reserved13 : Bool;   // Reserved
      reserved14 : Bool;   // Reserved
      reserved15 : Bool;   // Reserved
   END_STRUCT;
END_TYPE

TYPE "LIOLink_3RR24_typeMeasure"
TITLE = LIOLink_3RR24_typeMeasure
VERSION : 0.1
// Data set (index) 94 (measured values)
   STRUCT
      reserved : Array[0..15] of Byte;   // Reserve 0 - E-8 Dataset Index 94 Page 208
      activeCurrentL1 : Word;   // Active current L1
      activeCurrentL2 : Word;   // Active current L2
      activeCurrentL3 : Word;   // Active current L3
      activeCurrentMin : Word;   // Active current min
      activeCurrentMax : Word;   // Active current max
      activeCurrentAvg : Word;   // Active current avg
      apparentCurrentL1 : Word;   // Apparent current L1
      apparentCurrentL2 : Word;   // Apparent current L2
      apparentCurrentL3 : Word;   // Apparent current L3
      apparentCurrentMin : Word;   // Apparent current min
      apparentCurrentMax : Word;   // Apparent current max
      apparentCurrentAvg : Word;   // Apparent current avg
      activeVoltage : Word;   // Active voltage
      cosinePhi : Word;   // Cos phi value
      asymmetrySiemens : Word;   // Asymmetry Siemens
      asymmetryIecNema : Word;   // Asymmetry IEC/NEMA
      switchCounter : DWord;   // Switching cycle counter
      runtimeMeter : DWord;   // Runtime meter
   END_STRUCT;
END_TYPE

TYPE "LIOLink_3RR24_typeParam"
TITLE = LIOLink_3RR24_typeParam
VERSION : 0.1
// Data set (index) 131 (parameters)
   STRUCT
      reserved : Array[0..15] of Byte;   // Reserved
      groupDiagnostics : Bool := TRUE;   // Group diagnostics: Default: true, false; disabled, true: enabled
      groupErrorDiagnostics : Bool := TRUE;   // Group error diagnostics: Default: true, false; disabled, true: enabled
      reserved1 : Bool;   // Reserved
      reserved2 : Bool;   // Reserved
      localLimitChange : Bool := TRUE;   // Local threshold change: Default: true, false; disabled, true: enabled
      localParameterChange : Bool := TRUE;   // Local parameter change: Default: true, false; disabled, true: enabled
      localReset : Bool := TRUE;   // Local reset: Default: true, false; disabled, true: enabled
      retentiveErrorMemory : Bool;   // Retentitve error memory: Default: false, false; disabled, true: enabled
      analogValueCoding : Byte := 16#14;   // Analog value coding: Default: 20, Min: 0 (disabled), Max: 255
      reserved3 : Array[18..23] of Byte;   // Reserved
      resetResponse : Byte := 16#01;   // Reset response: Default: true, false: manual, true: automatic
      delayTimePowerOn : Bool := TRUE;   // ON-delay time (at Power ON): Default: true, false: disabled, true: enabled
      delayTimePowerOn0 : Bool;   // False
      delayTimeManResetOn : Bool := TRUE;   // ON-delay time (at manual reset): Default: true, false; disabled, true: enabled
      delayTimeManResetOn0 : Bool;   // False
      delayTimeRestartOn : Bool := TRUE;   // ON-delay time (at restart): Default: true, false; disabled, true: enabled
      delayTimeRestartOn0 : Bool;   // False
      reserved4 : Bool;   // Reserved
      reserved5 : Bool;   // Reserved
      phaseFault : Bool := TRUE;   // Phase failure monitoring: Default: true, false; disabled, true: enabled
      phaseFault0 : Bool;   // False
      phaseSequence : Bool := FALSE;   // Phase sequence monitoring: Default: false, false; disabled, true: enabled
      phaseSequence0 : Bool;   // False
      loadCurrent : Bool := FALSE;   // Load current monitoring(apparent current Is/active current Ip): Default: false, false: Is, true: Ip
      loadCurrent0 : Bool;   // False
      faultcurrent : Bool := FALSE;   // Fault current monitoring: Default: false, false; disabled, true: enabled
      faultcurrent0 : Bool;   // False
      asymmetry : Byte := 16#00;   // Asymmetry algorithm: Default: 0, 0: Siemens 1:IEC/NEMA
      delayTimeOn : Word := 16#0000;   // ON-delay time: Resolution: 0.1s=1, Default: 0s, Min: 0.1s or 0s (disabled), Max: 999,9s
      delayTimeTripUp : Word := 16#0000;   // Tripping delay time(current overshoot): Resolution: 0.1s=1, Default: 0s, Min: 0.1s or 0s (disabled), Max: 999,9s
      delayTimeTripDown : Word := 16#0000;   // Tripping delay time(current undrshoot): Resolution: 0.1s=1, Default: 0s, Min: 0.1s or 0s (disabled), Max: 999,9s
      delayTimeTripAsymmetry : Word := 16#0000;   // Tripping delay time(current asymmetry): Resolution: 0.1s=1, Default: 0s, Min: 0.1s or 0s (disabled), Max: 999,9s
      delayTimeReclose : Word := 16#0000;   // Reclosing delay time: Resolution: 0.1min=1, Default: 0min ,Min: 0.1min or 0min, Max: 300 min
      tresholdUp : Word := 16#0000;   // Threshold overshoot: 3RR2441(S00): Min: 1.6,Max: 16A ; 3RR2442(S0): Min: 4.0, Max: 40A
      tresholdDown : Word := 16#0000;   // Threshold undershoot: 3RR2441(S00): Min: 1.6, Max: 16A; 3RR2442(S0): Min: 4,0, Max: 40A
      tresholdAsymmetry : Word := 16#0000;   // Threshold current asymmetry: Resolution: 0.1%=1, Default: 0, Min: 5%, Max: 50%
      warningTresholdUp : Word := 16#0000;   // Warning threshold overshoot: 3RR2441(S00): Min: 1.6, Max: 16A; 3RR2442(S0): Min: 4.0, Max: 40A
      warningTresholdDown : Word := 16#0000;   // Warning threshold undershoot: 3RR2441(S00): Min:1.6, Max: 16A; 3RR2442(S0): Min: 4.0, Max: 40A
      warningTresholdAsymmetry : Word := 16#0000;   // Warning threshold current asymmetry: Resloution: 0.1%=1, Default: 0, Min: 5%, Max: 50%
      reserved6 : Array[50..55] of Byte;   // Reserved
      hysteresis : Word := 16#0000;   // Hysteresis (current): 3RR2441(S00): Min: 0.1, Max: 3A; 3RR2442(S0): Min:0.1, Max: 8A
      blockMonitoring : Word := 16#0000;   // Blocking current monitoring: Default: 0, Min: 2 or 0 (disabled), Max: 5
      reserved7 : Byte;   // Reserved
      relaySwitchResponse : Byte;   // Relay switching response:Default: 16#00, 16#00: Closed-circuit (NC), 16#01: Open-circuit(NO)
   END_STRUCT;
END_TYPE

TYPE "LIOLink_3RR24_typeAll"
TITLE = LIOLink_3RR24_typeAll
VERSION : 0.1
// Contains all the information about 3RR24
   STRUCT
      parameterPage0 : "LIOLink_typeParameterPage0";   // ID0: Parameter page 0
      systemCommands : Byte;   // ID2: System Commands (0x80 for device reset, 0x82 for factory reset, 0xA0 for switching cycle counter reset, 0xA1 for runtime meter reset) / ID2: Systemkommandos (0x80 für Device Reset, 0x82 für Factory Reset, 0xA0 für Schaltspielzähler Reset, 0xA1 für Betriebsstundenzähler Reset)
      vendorName : String[11];   // ID16: Vendor name / ID16: Herstellername
      vendorText : String[64];   // ID17: Vendor text / ID17: Herstellertext
      productName : String[64];   // ID18: Product name / ID18: Produktname
      productID : String[14];   // ID19: Product ID / ID19: Produkt ID
      serialNumber : String[16];   // ID21: Serial number / ID21: Seriennummer
      hwRevision : String[7];   // ID22: Hardware revision / ID22: Hardwarerevision
      fwRevision : String[7];   // ID23: Firmware revision / ID23: Firmwarerevision
      appSpecificName : String[32];   // ID24: Application specific name / ID24: Spezifischer Applikationsname
      diagnostics : "LIOLink_3RR24_typeDiag";   // ID92: Diagnostics / ID92: Diagnose
      measuredValues : "LIOLink_3RR24_typeMeasure";   // ID94: Measurement values / ID94: Messwerte
      parameters : "LIOLink_3RR24_typeParam";   // ID131: Parameters / ID131: Parameter
   END_STRUCT;
END_TYPE

// folder: LIOLink/Common/Device-specific data types/SIRIUS/3RS1

TYPE "LIOLink_3RS1_typeMeasure"
TITLE = LIOLink_3RS1_typeMeasure
VERSION : 0.1
// Data set (index) 94 (measured values)
   STRUCT
      reserved : Array[0..15] of Byte;   // Reserved
      sensorTemp1C : Int;   // Temperature in °C (Temperature sensor 1)
      sensorTemp1F : Int;   // Temperature in °F (Temperature sensor 1)
      sensorTemp2C : Int;   // Temperature in °C (Temperature sensor 2)(TEMP. 2 3RS1441 ONLY)
      sensorTemp2F : Int;   // Temperature in °F (Temperature sensor 2)(TEMP. 2 3RS1441 ONLY)
      sensorTemp3C : Int;   // Temperature in °C (Temperature sensor 3)(TEMP. 3 3RS1441 ONLY)
      sensorTemp3F : Int;   // Temperature in °F (Temperature sensor 3)(TEMP. 3 3RS1441 ONLY)
      tempMinC : Int;   // Temperature Tmin in °C
      tempMinF : Int;   // Temperature Tmin in °F
      tempMaxC : Int;   // Temperature Tmax in °C
      tempMaxF : Int;   // Temperature Tmax in °F
      tempAvgC : Int;   // Temperature Tavg in °C
      tempAvgF : Int;   // Temperature Tavg in °F
      reserved1 : Array[40..45] of Byte;   // Reserved
   END_STRUCT;
END_TYPE

TYPE "LIOLink_3RS1_typeParam"
TITLE = LIOLink_3RS1_typeParam
VERSION : 0.1
// Data set (index) 131 - parameters
   STRUCT
      reserved : Array[0..15] of Byte;   // Reserved
      groupDiagnostic : Bool := TRUE;   // Group diagnostics: Default: True, False: disabled, True: enabled
      groupError : Bool := TRUE;   // Group error diagnostics: Default: True, False: disabled, True: enabled
      reserved1 : Bool;   // Reserved
      reserved2 : Bool;   // Reserved
      localLimitChange : Bool := TRUE;   // Local threshold change: Default: True, False: disabled, True: enabled
      localParamChange : Bool := TRUE;   // Local parameter change: Default: True, False: disabled, True: enabled
      localReset : Bool := TRUE;   // Local reset: Default: True, False: disabled, True: enabled
      retentiveErrorMem : Bool := FALSE;   // Retentive error memory: Default: False, False: disabled, True: enabled
      analogValueCoding : USInt := 5;   // Analog value coding: Default: 5, Min: 0 (disabled), Max: 255
      reserved3 : Array[18..23] of Byte;   // Reserved
      reserved4 : Bool;   // Reserved
      reserved5 : Bool;   // Reserved
      monitorMode1 : Bool := FALSE;   // Temp. monitoring mode:Default: False, False: Overshoot/Range Monitor, True: Undershoot
      monitorMode2 : Bool := FALSE;   // Temp. monitoring mode:Default: False, False: Overshoot/Undershoot , True: Range Monitor
      monitorMode3 : Bool := FALSE;   // False
      unit : Bool;   // Temperature unit: False:°C (degrees Celcius) True:°F (degrees Fahrenheit)
      unit0 : Bool := FALSE;   // False
      unit1 : Bool;   // False
      delayOn : Bool := TRUE;   // ON-delay time (at Power ON): Default: true, false: disabled, true: enabled
      delayOn0 : Bool;   // False
      delayManual : Bool := TRUE;   // ON-delay time (at manual reset): Default: true, false: disabled, true: enabled
      delayManual0 : Bool;   // False
      reserved6 : Bool;   // Reserved
      reserved7 : Bool;   // Reserved
      reserved8 : Bool;   // Reserved
      reserved9 : Bool;   // Reserved
      delayTimeOn : Int;   // ON-delay time: Resolution:0,1s=1,Default:0,Min:1 or 0(disabled),Max:999,9s
      delayTimeLevel : Int;   // Tripping delay time(temp.ovr-/undrsht):Rsltn:0,1s=1,Dflt:0,Min:1or.0,Max:999,9s
      reserved10 : Byte;   // Reserved
      sensor1Available : Bool := TRUE;   // 3RS1440/3RS1441/3RS1540:Temperature sensor 1: False: disabled, true: enabled
      sensor2Available : Bool;   // 3RS1441 ONLY: Temperature sensor 2: False: disabled, true: enabled, Default: true
      sensor3Available : Bool;   // 3RS1441 ONLY: Temperature sensor 3: False: disabled, true: enabled, Default: true
      reserved11 : Bool;   // Reserved
      reserved12 : Bool;   // Reserved
      reserved13 : Bool;   // Reserved
      reserved14 : Bool;   // Reserved
      reserved15 : Bool;   // Reserved
      sensorType : USInt;   // Temperature sensor type: 3RS1440/1441 resistance sensor, 3RS1540 thermocouple
      limitValueV1 : Int := 80;   // Limit value v1: Min:-50(resist.sensors)/-99°(thermocouples)C, Max:750/1800°C
      limitValueV2 : Int := 50;   // Limit value v2: Min:-50(resist.sensors)/-99°C(thermocouples), Max:750/1800°C
      warningValueV1 : Int := 72;   // Warning threshold v1: Min:-50(resist.sen.)/-99°C(thermocouples), Max:750/1800°C
      warningValueV2 : Int := 45;   // Warning threshold v2: Min:-50(resist.sen.)/-99°C(thermocouples), Max:750/1800°C
      reserved16 : Array[42..45] of Byte;   // Reserved
      hysteresis : Word := 16#0005;   // Hysteresis: Default: 5°C/5°F, Min:1°C/1°F or 0 (disabled),Max:99°C/99°F
      relaySwitchResponse : Bool := FALSE;   // Relay switching response:Default: false, false: Closed-circuit(NC), true: Open-ciruict(NO)
      relaySwitchResponse0 : Bool;   // False
      reserved17 : Bool;   // Reserved
      reserved18 : Bool;   // Reserved
      reserved19 : Bool;   // Reserved
      reserved20 : Bool;   // Reserved
      reserved21 : Bool;   // Reserved
      reserved22 : Bool;   // Reserved
      reserved23 : Byte;   // Reserved
   END_STRUCT;
END_TYPE

TYPE "LIOLink_3RS1_typeSensor"
TITLE = LIOLink_3RS1_typeSensor
// Temperature monitoring, part of the data set (index) 92 - diagnostics
   STRUCT
      rangeOvershoot : Bool;   // Temperature sensor - Measuring range overshoot
      wireBreak : Bool;   // Temperature sensor - Wire break
      shortCircuit : Bool;   // Temperature sensor - Short-circuit
      reserved13 : Bool;   // Reserved
      reserved14 : Bool;   // Reserved
      reserved15 : Bool;   // Reserved
      reserved16 : Bool;   // Reserved
      reserved17 : Bool;   // Reserved
      aboveBothLimits : Bool;   // Temperature sensor - Measured value above the two limit values (overshoot)
      aboveFirstLimit : Bool;   // Temperature sensor - Measured value above first limit value (overshoot)
      withinRange : Bool;   // Temperature sensor - Measured value within range of limit values
      belowFirstLimit : Bool;   // Temperature sensor - Measured value below first limit value (undershoot)
      belowBothLimits : Bool;   // Temperature sensor - Measured value below the two limit values (undershoot)
      reserved18 : Bool;   // Reserved
      reserved19 : Bool;   // Reserved
      reserved20 : Bool;   // Reserved
      aboveBothWarningLimits : Bool;   // Temperature sensor - Measured value above two warning thresholds (overshoot)
      aboveFirstWarningLimit : Bool;   // Temperature sensor - Measured value above first warning threshold (overshoot)
      withinRangeWarning : Bool;   // Temperature sensor - Measured value within range of warning threshold
      belowFirstWarningLimit : Bool;   // Temperature sensor - Measured value below first warning threshold (undershoot
      belowBothWarningLimits : Bool;   // Temperature sensor - Measured value below two warning threshold (undershoot)
      reserved21 : Bool;   // Reserved
      reserved22 : Bool;   // Reserved
      reserved23 : Bool;   // Reserved
      reserved24 : Byte;   // Reserved
   END_STRUCT;
END_TYPE

TYPE "LIOLink_3RS1_typeDiag"
TITLE = LIOLink_3RS1_typeDiag
VERSION : 0.1
// Data set (index) 92 - diagnostics
   STRUCT
      reserved : Array[0..15] of Byte;   // Reserved
      ready : Bool;   // Ready
      groupError : Bool;   // Group error
      generalWarning : Bool;   // General warning
      reserved1 : Bool;   // Reserved
      reserved2 : Bool;   // Reserved
      parameterAssign : Bool;   // Parameter assignment active
      parameterInvalid : Bool;   // Invalid parameter
      internalError : Bool;   // Self-test error/internal error
      reserved3 : Bool;   // Reserved
      errorNumber : Word;   // Parameter error number
      reserved4 : Array[20..25] of Byte;   // Reserved
      delayTimeRunning : Bool;   // ON-delay time running
      delayLevelUp : Bool;   // Tripping delay time running (limit value v1 or limit value v2)
      reserved5 : Bool;   // Reserved
      reserved6 : Bool;   // Reserved
      reserved7 : Bool;   // Reserved
      reserved8 : Bool;   // Reserved
      reserved9 : Bool;   // Reserved
      reserved10 : Bool;   // Reserved
      levelV1Up : Bool;   // Limit value v1 overshoot
      levelV2Up : Bool;   // Limit value v2 overshot
      levelV1UpWarning : Bool;   // Warning limit for v1 overshoot
      levelV2UpWarning : Bool;   // Warning limit for v2 overshoot
      resetResponse : Bool;   // Reset response:0:Manual reset,1:Autorst/permanent jmpr between terminals y3/y4
      reserved11 : Bool;   // Reserved
      reserved12 : Bool;   // Reserved
      reserved13 : Bool;   // Reserved
      sensor : Array[1..3] of "LIOLink_3RS1_typeSensor";   // Temperature monitoring
   END_STRUCT;
END_TYPE

TYPE "LIOLink_3RS1_typeAll"
TITLE = LIOLink_3RS1_typeAll
VERSION : 0.1
// Contains all the information about 3RS1
   STRUCT
      parameterPage0 : "LIOLink_typeParameterPage0";   // ID0: Parameter page 0
      vendorName : String[11];   // ID16: Vendor name / ID16: Herstellername
      vendorText : String[64];   // ID17: Vendor text / ID17: Herstellertext
      productName : String[64];   // ID18: Product name / ID18: Produktname
      productID : String[14];   // ID19: Product ID / ID19: Produkt ID
      hardwareRevision : String[7];   // ID22: Hardware revision / ID22: Hardwarerevision
      firmwareRevision : String[7];   // ID23: Firmware revision / ID23: Firmwarerevision
      appSpecificName : String[32];   // ID24: Application specific name / ID24: Spezifischer Applikationsname
      diagnostics : "LIOLink_3RS1_typeDiag";   // ID92: Diagnostics / ID92: Diagnose
      measuredValues : "LIOLink_3RS1_typeMeasure";   // ID94: Measurement values / ID94: Messwerte
      parameters : "LIOLink_3RS1_typeParam";   // ID131: Parameters / ID131: Parameter
   END_STRUCT;
END_TYPE

// folder: LIOLink/Common/Device-specific data types/SIRIUS/3RS2

TYPE "LIOLink_3RS2_typeCurrentInput"
TITLE = LIOLink_3RS2_typeCurrentInput
// Part of the Data set 92 - Diagnostics, Current Input 4..20mA
   STRUCT
      overstepping : Bool;   // Measuring range overstepping
      res0 : Bool;   // Reserved
      res1 : Bool;   // Reserved
      res2 : Bool;   // Reserved
      res3 : Bool;   // Reserved
      res4 : Bool;   // Reserved
      res5 : Bool;   // Reserved
      res6 : Bool;   // Reserved
      aboveBothLimits : Bool;   // Measured value is above the two limit values (monitoring for overshoot)
      aboveFirstLimit : Bool;   // Measured value is above the first limit value (monitoring for overshoot)
      withinRangeLimits : Bool;   // Measured value is within range of limit values
      belowFirstLimit : Bool;   // Measured value is below the first limit value for overshoot (monitoring for undershoot)
      belowBothLimits : Bool;   // Measured value is below the two limit values (monitoring for undershoot)
      res7 : Bool;   // Reserved
      res8 : Bool;   // Reserved
      res9 : Bool;   // Reserved
      aboveBothWarningLimits : Bool;   // Measured value is above the two warning limits (monitoring for overshoot)
      aboveFirstWarningLimit : Bool;   // Measured value is above the first warning limit (monitoring for overshoot)
      withinRangeWarningLimits : Bool;   // Measured value is within range of warning limits
      belowFirstWarningLimit : Bool;   // Measured value is below the first warning limit for overshoot (monitoring for undershoot)
      belowBothWarningLimits : Bool;   // Measured value is below the two warning limits (monitoring for undershoot)
      res10 : Bool;   // Reserved
      res11 : Bool;   // Reserved
      res12 : Bool;   // Reserved
      res13 : Byte;   // Reserved
   END_STRUCT;
END_TYPE

TYPE "LIOLink_3RS2_typeMeasureFloat"
TITLE = LIOLink_3RS2_typeMeasureFloat
// Data set 95 - measured values (floating-point format)
   STRUCT
      reserved : Array[0..15] of Byte;   // Reserved
      sensorTemp1C : Real;   // Temperature in °C (Temperature sensor 1)
      sensorTemp1F : Real;   // Temperature in °F (Temperature sensor 1)
      sensorTemp2C : Real;   // Temperature in °C (Temperature sensor 2)
      sensorTemp2F : Real;   // Temperature in °F (Temperature sensor 2)
      sensorTemp3C : Real;   // Temperature in °C (Temperature sensor 3)
      sensorTemp3F : Real;   // Temperature in °F (Temperature sensor 3)
      tempMinC : Real;   // Temperature Tmin in °C
      tempMinF : Real;   // Temperature Tmin in °F
      tempMaxC : Real;   // Temperature Tmax in °C
      tempMaxF : Real;   // Temperature Tmax in °F
      tempAvgC : Real;   // Temperature Tavg in °C
      tempAvgF : Real;   // Temperature Tavg in °F
      currentInput : Real;   // Current input
   END_STRUCT;
END_TYPE

TYPE "LIOLink_3RS2_typeSensor"
TITLE = LIOLink_3RS2_typeSensor
// Part of Data set 92 - Diagnostics, diagnostics of sensor
   STRUCT
      rangeOvershoot : Bool;   // Measuring range overshoot
      wireBreak : Bool;   // Wire break
      shortCircuit : Bool;   // Short-circuit
      reserved : Bool;   // Reserved
      reserved1 : Bool;   // Reserved
      reserved2 : Bool;   // Reserved
      reserved3 : Bool;   // Reserved
      reserved4 : Bool;   // Reserved
      aboveBothLimits : Bool;   // Measured value is above the two limit values (monitoring for overshoot)
      aboveFirstLimit : Bool;   // Measured value is above the first limit value (monitoring for overshoot)
      withinRange : Bool;   // Measured value is within range of limit values
      belowFirstLimit : Bool;   // Measured value is below the first limit value for overshoot (monitoring for undershoot)
      belowBothLimits : Bool;   // Measured value is below the two limit values (monitoring for undershoot)
      reserved5 : Bool;   // Reserved
      reserved6 : Bool;   // Reserved
      reserved7 : Bool;   // Reserved
      aboveBothWarningLimits : Bool;   // Measured value is above the two warning limits (monitoring for overshoot)
      aboveFirstWarningLimit : Bool;   // Measured value is above the first warning limit (monitoring for overshoot)
      withinRangeWarning : Bool;   // Measured value is within range of warning limits
      belowFirstWarningLimit : Bool;   // Measured value is below the first warning limit for overshoot (monitoring for undershoot)
      belowBothWarningLimits : Bool;   // Measured value is below the two warning limits (monitoring for undershoot)
      reserved8 : Bool;   // Reserved
      reserved9 : Bool;   // Reserved
      reserved10 : Bool;   // Reserved
      reserved11 : Byte;   // Reserved
   END_STRUCT;
END_TYPE

TYPE "LIOLink_3RS2_typeMeasure"
TITLE = LIOLink_3RS2_typeMeasure
VERSION : 0.1
// Data set 94 - measured values
   STRUCT
      reserved : Array[0..15] of Byte;   // Reserved
      sensorTemp1C : Int;   // Temperature in °C (Temperature sensor 1)
      sensorTemp1F : Int;   // Temperature in °F (Temperature sensor 1)
      sensorTemp2C : Int;   // Temperature in °C (Temperature sensor 2)
      sensorTemp2F : Int;   // Temperature in °F (Temperature sensor 2)
      sensorTemp3C : Int;   // Temperature in °C (Temperature sensor 3)
      sensorTemp3F : Int;   // Temperature in °F (Temperature sensor 3)
      tempMinC : Int;   // Temperature Tmin in °C
      tempMinF : Int;   // Temperature Tmin in °F
      tempMaxC : Int;   // Temperature Tmax in °C
      tempMaxF : Int;   // Temperature Tmax in °F
      tempAvgC : Int;   // Temperature Tavg in °C
      tempAvgF : Int;   // Temperature Tavg in °F
      currentInput : Int;   // Current input
   END_STRUCT;
END_TYPE

TYPE "LIOLink_3RS2_typeParam"
TITLE = LIOLink_3RS2_typeParam
VERSION : 0.1
// Data set 131 - parameters
   STRUCT
      reserved : Array[0..15] of Byte;   // Reserved
      groupDiag : Bool := TRUE;   // Group diagnostics: Default: True, False: disabled, True: enabled
      groupErrorDiag : Bool := TRUE;   // Group error diagnostics: Default: True, False: disabled, True: enabled
      reserved1 : Bool;   // Reserved
      reserved2 : Bool;   // Reserved
      localLimChange : Bool := TRUE;   // Local limit change: Default: True, False: disabled, True: enabled
      localParamChange : Bool := TRUE;   // Local parameter change: Default: True, False: disabled, True: enabled
      localReset : Bool := TRUE;   // Local reset: Default: True, False: disabled, True: enabled
      retentiveErrorMem : Bool := TRUE;   // Retentive error memory: Default: True, False: disabled, True: enabled
      analogValueCoding : USInt := 5;   // Analog value coding: Default: 5, Min: 1, Max: 160
      reserved3 : Array[18..23] of Byte;   // Reserved
      reset : Bool;   // Reset: Default: False, False: manual, True: auto
      reserved5 : Bool;   // Reserved
      monitorMode1 : Bool;   // Monitoring mode [0] overshoot [Default]; [1] undershoot; [2] window monitoring
      monitorMode2 : Bool;   // Monitoring mode [0] overshoot [Default]; [1] undershoot; [2] window monitoring
      monitorMode3 : Bool;   // Monitoring mode [0] overshoot [Default]; [1] undershoot; [2] window monitoring
      unit1 : Bool;   // Temperature unit [0]°C [Default]; [1] °F; [2] mA; [3] %
      unit2 : Bool;   // Temperature unit [0]°C [Default]; [1] °F; [2] mA; [3] %
      unit3 : Bool;   // Temperature unit [0]°C [Default]; [1] °F; [2] mA; [3] %
      onDelayStart : Bool;   // ON-delay time (at Power ON): Default: [0], [0] disabled, [1] enabled
      reserved6 : Bool;   // Reserved
      onDelayReset : Bool;   // ON-delay time (at manual reset): Default: [0], [0] disabled, [1] enabled
      reserved7 : Bool;   // Reserved
      reserved8 : Bool;   // Reserved
      reserved9 : Bool;   // Reserved
      reserved10 : Bool;   // Reserved
      reserved11 : Bool;   // Reserved
      startupDly : Int;   // Startup delay; Resolution: 0.1s=1, Default: 0, Min: 1 or 0 (disabled), Max: 9999 * 0.1 s = 999.9 s
      tripDly : Int;   // Tripping delay time (if the temperature is overshot or undershot); Resolution: 0.1s=1, Default: 0, Min: 1 or 0 (disabled), Max: 9999 * 0.1 s = 999.9 s
      reserved12 : Int;   // Reserved
      sensor1En : Bool := TRUE;   // Sensor 1 enabled; Default: False, False: disabled, True: enabled
      sensor2En : Bool;   // Sensor 2 enabled; Default: False, False: disabled, True: enabled
      sensor3En : Bool;   // Sensor 3 enabled; Default: False, False: disabled, True: enabled
      currentInputEn : Bool;   // Current input 4..20 mA enabled; Default: False, False: disabled, True enabled
      sensorExpModule : Bool;   // Sensor expansion module / output relay K3; Default: False, False: disabled, True enabled
      reserved13 : Bool;   // Reserved
      reserved14 : Bool;   // Reserved
      reserved15 : Bool;   // Reserved
      sensorType : Byte := 16#80;   // Sensor type; Default: 128, 128: Pt100 (2-wire), 129: Pt1000 (2-wire), 130: KTY83 (2-wire), 131: KTY84 (2-wire), 132: NTC (2-wire), 136: Pt100 (3-wire), 137: Pt1000 (3-wire), 138: KTY83 (3-wire), 139: KTY84 (3-wire), 140: NTC (3-wire), 1: J, 2: K, 3: T, 4: E, 5: N, 6: S, 7: R, 8: B, 160: current input 4..20 mA
      limitV1 : Int := 80;   // Limit v1; Default: 80, Min: -50 °C (resistance sensors) / -99 °C (thermocouples), Max: 750 °C (resistance sensors)/1800 °C (thermocouples)
      limitV2 : Int := 50;   // Limit v2; Default: 50, Min: -50 °C (resistance sensors) / -99 °C (thermocouples), Max: 750 °C (resistance sensors)/1800 °C (thermocouples)
      warnLimitV1 : Int := 75;   // Warning limit v1; Default: 75, Min: -50 °C (resistance sensors) / -99 °C (thermocouples), Max: 750 °C (resistance sensors)/1800 °C (thermocouples)
      warnLimitV2 : Int := 45;   // Warning limit v2; Default: 45, Min: -50 °C (resistance sensors) / -99 °C (thermocouples), Max: 750 °C (resistance sensors)/1800 °C (thermocouples)
      reserved16 : DWord;   // Reserved
      hysteresis : Int := 5;   // Hysteresis; Default: 5 °C / 5 °F, Min: 1 °C/1 °F, Max: 999 °C / 999 °F
      relayBehavior : Bool;   // Relay switching behavior; Default: False, False: Quiescent current principle, True Open-circuit principle
      reserved17 : Bool;   // Reserved
      reserved18 : Bool;   // Reserved
      reserved19 : Bool;   // Reserved
      reserved20 : Bool;   // Reserved
      reserved21 : Bool;   // Reserved
      reserved22 : Bool;   // Reserved
      reserved23 : Bool;   // Reserved
      reserved24 : Byte;   // Reserved
      minRange : Int := 40;   // Current input 4..20 mA minimum range; Default: 40, Min: -200 (°C/°F) / 0 (%), Max: 9999 (°C/°F) / 150 (%)
      maxRange : Int := 80;   // Current input 4..20 mA maximum range; Default: 40, Min: -200 (°C/°F) / 0 (%), Max: 9999 (°C/°F) / 150 (%)
      offsetSensor1 : Int;   // Offset sensor 1; Default: 0, Min: -99, Max: 99
      offsetSensor2 : Int;   // Offset sensor 2; Default: 0, Min: -99, Max: 99
      offsetSensor3 : Int;   // Offset sensor 3; Default: 0, Min: -99, Max: 99
      offsetCurrentInput : Int;   // Offset current input 4..20 mA; Default: 0, Min: -10.0 mA / -99 °C/°F, Max: 10.0 mA / 99 °C / °F, reading always returns 0
      compMeasuringPt : Int;   // Comparison measuring point in °C/°F; Default: 0, Min: -25 °C / -13 °F, Max: 80 °C / 176 °F, reading always returns 0
      ecoMode : Bool := TRUE;   // Eco mode; Default [1], [0] disabled, [1] enabled
      ponProtection : Bool;   // Pin Protection Default [0], [0] disabled, [1] enabled
      extCompMeasuringPt : Bool;   // External comparison measuring point; Default [0], [0] disabled, [1] enabled
      reserved25 : Bool;   // Reserved
      reserved26 : Bool;   // Reserved
      reserved27 : Bool;   // Reserved
      reserved28 : Bool;   // Reserved
      reserved29 : Bool;   // Reserved
      reserved30 : Byte;   // Reserved
      pin : Int;   // PIN; Default: 0, Min: 0, Max: 999, reading always returns 0
      newPin : Int;   // New PIN; Default: 0, Min: 0, Max: 999, reading always returns 0
      deviceMode : Byte;   // Device mode; Default: [0], [0] standard, [1] ATEX, [2] Temperature monitor TW, [3] Temperature limiter TB
      reserved31 : Byte;   // Reserved
   END_STRUCT;
END_TYPE

TYPE "LIOLink_3RS2_typeDiag"
TITLE = LIOLink_3RS2_typeDiag
VERSION : 0.1
// Data set 92 - Diagnostics
   STRUCT
      reserved : Array[0..15] of Byte;   // Reserved
      ready : Bool;   // Ready
      groupError : Bool;   // Group error
      groupWarning : Bool;   // Group warning
      reserved1 : Bool;   // Reserved
      communicationError : Bool;   // Sensor expansion module - communication error
      parameterAssign : Bool;   // Parameter assignment active
      parameterInvalid : Bool;   // Invalid parameter
      internalError : Bool;   // Self-test error/internal error
      paramAckReq : Bool;   // Parameter confirmation required
      reserved2 : Bool;   // Reserved
      reserved3 : Bool;   // Reserved
      reserved4 : Bool;   // Reserved
      reserved5 : Bool;   // Reserved
      reserved6 : Bool;   // Reserved
      reserved7 : Bool;   // Reserved
      reserved8 : Bool;   // Reserved
      errorNumber : Word;   // Incorrect parameter number
      reserved9 : Array[20..25] of Byte;   // Reserved
      delayTimeRunning : Bool;   // ON-delay time running
      delayLevelUpV1 : Bool;   // Tripping delay time running (limit value v1)
      delayLevelUpV2 : Bool;   // Tripping delay time running (limit value v2)
      reserved10 : Bool;   // Reserved
      reserved11 : Bool;   // Reserved
      reserved12 : Bool;   // Reserved
      reserved13 : Bool;   // Reserved
      reserved14 : Bool;   // Reserved
      levelV1UpDown : Bool;   // Limiting value v1 overshot/undershot
      levelV2UpDown : Bool;   // Limiting value v2 overshot/undershot
      levelV1Warning : Bool;   // Warning limit v1 overshot/undershot
      levelV2Warning : Bool;   // Warning limit v1 overshot/undershot
      reserved15 : Bool;   // Reserved
      reserved16 : Bool;   // Reserved
      reserved17 : Bool;   // Reserved
      reserved18 : Bool;   // Reserved
      sensor : Array[1..3] of "LIOLink_3RS2_typeSensor";   // Temperature sensor 1
      currentInput : "LIOLink_3RS2_typeCurrentInput";   // Current input
   END_STRUCT;
END_TYPE

TYPE "LIOLink_3RS2_typeAll"
TITLE = LIOLink_3RS2_typeAll
VERSION : 0.1
// Contains all the information about 3RS2
   STRUCT
      parameterPage0 : "LIOLink_typeParameterPage0";   // ID0: Parameter page 0
      systemCommand : Byte;   // ID2: System commands
      vendorName : String[11];   // ID16: Vendor name
      vendorText : String[64];   // ID17: Vendor text
      productName : String[64];   // ID18: Product name
      productID : String[14];   // ID19: Product ID
      firmwareRevision : String[7];   // ID23: Firmware revision
      appSpecificName : String[32];   // ID24: Application specific name
      diagnostics : "LIOLink_3RS2_typeDiag";   // ID92: Diagnostics
      measuredValues : "LIOLink_3RS2_typeMeasure";   // ID94: Measurement values
      measuredValuesFloat : "LIOLink_3RS2_typeMeasureFloat";   // ID95: Measurement as floating values
      parameters : "LIOLink_3RS2_typeParam";   // ID131: Parameters
   END_STRUCT;
END_TYPE

// folder: LIOLink/Common/Device-specific data types/SIRIUS/3SU1/3SU1 Electronic Module

TYPE "LIOLink_3SU1_ElecModule_typeAll"
TITLE = LIOLink_3SU1_ElecModule_typeAll
VERSION : 0.1
// Contains all the information about 3SU1 ElecModule
   STRUCT
      parameterPage0 : "LIOLink_typeParameterPage0";   // ID0: Parameter page 0
      systemCommand : Byte;   // Write System Command to Device: 0xA1 - 0xB1; 0x82 = Default
      vendorName : String[10];   // ID16: Vendor name
      vendorText : String[64];   // ID17: Vendor text
      productName : String[64];   // ID18: Product name
      productID : String[18];   // ID19: Product ID
      fwRevision : String[6];   // ID23: Firmware revision
      appSpecificName : String[32];   // ID24: Application specific name
      processDataOut : Array[0..5] of Byte;   // ID67: Process Data of outputs
      processDataIn : Array[0..5] of Byte;   // ID69: Process Data of inputs
      diagnostics : "LIOLink_3SU1_ElecModule_typeDiag92";   // ID92: Diagnostics
      statistics : "LIOLink_3SU1_ElecModule_typeDiag94";   // ID94: Statistics
      parameters : "LIOLink_3SU1_ElecModule_typeParam";   // ID131: Parameters
   END_STRUCT;
END_TYPE

TYPE "LIOLink_3SU1_ElecModule_typeDiag92"
TITLE = LIOLink_3SU1_ElecModule_typeDiag92
VERSION : 0.1
// Diagnostics - data set (index) 92
   STRUCT
      reserved : Array[0..15] of Byte;   // Reserved
      status : Byte;   // Status: 1 = Ready; 2 = Error
      switchOnDuraStatIO0_3 : Byte;   // Switch-on duration status: 0x00=Inactive; 0x01=running; 0x02=reached; 0x03=finished
      switchOnDuraStatIO4_7 : Byte;   // Switch-on duration status: 0x00=Inactive; 0x01=running; 0x02=reached; 0x03=finished
      dimStatusOutputQ0_3 : Byte;   // Dimming status: 0x00=Inactive; 0x01=running; 0x03=finished
      dimStatusOutputQ4_7 : Byte;   // Dimming status: 0x00=Inactive; 0x01=running; 0x03=finished
      switchCycleCntStatIO0_3 : Byte;   // Switching cycle counter status: 0x00=Inactive; 0x01=running; 0x02=reached; 0x03=finished
      switchCycleCntStatIO4_7 : Byte;   // Switching cycle counter status: 0x00=Inactive; 0x01=running; 0x02=reached; 0x03=finished
      reserved1 : Byte;   // Reserved
   END_STRUCT;
END_TYPE

TYPE "LIOLink_3SU1_ElecModule_typeParam"
TITLE = LIOLink_3SU1_ElecModule_typeParam
VERSION : 0.1
// Parameters - Data set (index) 131
   STRUCT
      reserved : Array[0..15] of Byte;   // Reserved
      functionModeIO : Array[0..7] of Byte;   // 0x01=Input; 0x02=Output; 0x03=PWM; 0x04=Dimming Output; 0x05=InputCounter; 0x06=OutputCounter; 0x07=TurnonTimeInput; 0x08=TurnonTimeOutput
      setupGroup : Byte;   // 0x00=individual; 0x01=all; 0x02=grouped // .x3:1 = enable data reset
      pwmFreqQ : Array[0..7] of Byte;   // Range: 1..255; 1 = 1Hz
      pwmDutyQ : Array[0..7] of Byte;   // Range: 10 - 90 %; 1 = 1%
      dimmingTimeQ : Array[0..7] of Byte;   // Range: 1 - 255; 1 = 0.1Hz
      inputDelay : Array[0..7] of Byte;   // Range: 3-255; 1 = 1ms
      inputTimeThreshold : Array[0..7] of DWord;   // Set threshold for tripping due to a value overshoot: 1 = 1s
      inputCounterThreshold : Array[0..7] of DWord;   // Set threshold for tripping due to a value overshoot
      inputCounterEdgeI0_3 : Byte;   // 0x00=no edge; 0x01=rising edge; 0x02=falling edge; 0x03=all edges
      inputCounterEdgeI4_7 : Byte;   // 0x00=no edge; 0x01=rising edge; 0x02=falling edge; 0x03=all edges
      inputInvertI0_7 : Byte;   // 0=not inverted; 1=inverted
      outputInvertQ0_7 : Byte;   // 0=not inverted; 1=inverted
      reserved1 : Byte;   // Reserved
   END_STRUCT;
END_TYPE

TYPE "LIOLink_3SU1_ElecModule_typeDiag94"
TITLE = LIOLink_3SU1_ElecModule_typeDiag94
VERSION : 0.1
// Diagnostics - data set (index) 94
   STRUCT
      reserved : Array[0..15] of Byte;   // Reserved
      switchOnDurationsIO : Array[0..7] of DWord;   // Switch-on duration in seconds
      switchCycCountersIO : Array[0..7] of DWord;   // Switching cycle counter
      inputValue : Byte;   // Input value
      outputValue : Byte;   // Output value
   END_STRUCT;
END_TYPE

// folder: LIOLink/Common/Device-specific data types/SIRIUS/3SU1/3SU1 ID Key Switch

TYPE "LIOLink_3SU1_IDKeySwitch_typeKeyList2"
TITLE = LIOLink_3SU1_IDKeySwitch_typeKeyList2
VERSION : 0.1
// Data record (index) 82 - memory of the individually codable ID keys
   STRUCT
      keys : Array[31..50] of "LIOLink_3SU1_IDKeySwitch_typeKeyState";   // Data record (index) 82 - memory of the individually codable ID keys
   END_STRUCT;
END_TYPE

TYPE "LIOLink_3SU1_IDKeySwitch_typeDiag94"
TITLE = LIOLink_3SU1_IDKeySwitch_typeDiag94
VERSION : 0.1
// Data record (index) 94 (ID key)
   STRUCT
      reserved : Array[0..15] of Byte;   // Reserved
      insertedKey : "LIOLink_3SU1_IDKeySwitch_typeKeyState";   // Inserted ID key
   END_STRUCT;
END_TYPE

TYPE "LIOLink_3SU1_IDKeySwitch_typeDiag92"
TITLE = LIOLink_3SU1_IDKeySwitch_typeDiag92
VERSION : 0.1
// Data record (index) 92 - diagnostics
   STRUCT
      reserved : Array[0..15] of Byte;   // Reserved
      status : Byte;   // Status: 1 = Ready; 2 = Error
      outputs : Byte;   // Output state: Permission= .X0 - .X3 Key inserted= .X4
      detectionKey : Byte;   // Detection of the ID key
      statusKey : Byte;   // Status of the individually encodable ID Key
   END_STRUCT;
END_TYPE

TYPE "LIOLink_3SU1_IDKeySwitch_typeAll"
TITLE = LIOLink_3SU1_IDKeySwitch_typeAll
VERSION : 0.1
// Contains all the information about 3SU1 IDKeySwitch
   STRUCT
      parameterPage0 : "LIOLink_typeParameterPage0";   // ID0: Parameter page 0
      systemCommand : Byte;   // Write System Command to Device: 0xA1 - 0xA7; 0x82 = Default
      vendorName : String[10];   // ID16: Vendor name
      vendorText : String[64];   // ID17: Vendor text
      productName : String[64];   // ID18: Product name
      productID : String[18];   // ID19: Product ID
      fwRevision : String[5];   // ID23: Firmware revision
      appSpecificName : String[32];   // ID24: Application specific name
      processDataIn : Array[0..5] of Byte;   // ID69: Process data of inputs
      addKeyID : "LIOLink_3SU1_IDKeySwitch_typeKeyState";   // ID79: Add individually encodeable ID key
      delKeyID : "LIOLink_3SU1_IDKeySwitch_typeKeyState";   // ID80: Delete Individually encodeable ID key
      keyList1 : "LIOLink_3SU1_IDKeySwitch_typeKeyList1";   // ID81: List of saved indivually encodeable ID keys 1 to 30
      keyList2 : "LIOLink_3SU1_IDKeySwitch_typeKeyList2";   // ID82: List of saved indivually encodeable ID keys 31..50
      diagnostics : "LIOLink_3SU1_IDKeySwitch_typeDiag92";   // ID92: Diagnostics
      insertedKey : "LIOLink_3SU1_IDKeySwitch_typeDiag94";   // ID94: Inserted ID key
      parameters : "LIOLink_3SU1_IDKeySwitch_typeParam";   // ID131: Parameters
   END_STRUCT;
END_TYPE

TYPE "LIOLink_3SU1_IDKeySwitch_typeKeyList1"
TITLE = LIOLink_3SU1_IDKeySwitch_typeKeyList1
VERSION : 0.1
// Data record (index) 81 - memory of the individually codable ID keys
   STRUCT
      keys : Array[1..30] of "LIOLink_3SU1_IDKeySwitch_typeKeyState";   // Data record (index) 81 - memory of the individually codable ID keys
   END_STRUCT;
END_TYPE

TYPE "LIOLink_3SU1_IDKeySwitch_typeParam"
TITLE = LIOLink_3SU1_IDKeySwitch_typeParam
VERSION : 0.1
// Data record (index) 131 (parameters)
   STRUCT
      reserved : Array[0..15] of Byte;   // Reserved
      switchInStages : Bool;   // Switch in stages; 0: disabled, 1: enabled
      switchPosMemory : Bool;   // Switch position memory; 0: disabled (key position = 0), 1: enabled (last key position is retained)
      switchPosRetentive : Bool;   // Switch position retentive memory; 0: disabled, 1: enabled
      individualOnly : Bool;   // Individually encodeable ID keys only; 0: disabled, 1: enabled
      reserved1 : Bool;   // Reserved
      reserved2 : Bool;   // Reserved
      reserved3 : Bool;   // Reserved
      reserved4 : Bool;   // Reserved
      switchPosDelay : Byte;   // Switch position delay; 1 = 0.1 s (0 to 100)
      selectMem : Byte;   // Select memory range (1 to 5)
      deactSwitchOff : Bool;   // Deactivation of switch-off function (>= V2.0.0)
      deactRedLed : Bool;   // Deactivate red LEDs (>= V2.0.0)
      reductAuthLevel : Bool;   // Permit a reduction of the authorization level via the switch (>= V2.0.0)
      actLampTest : Bool;   // Activate lamp test (>= V2.0.0)
      reserved5 : Bool;   // Reserved
      reserved6 : Bool;   // Reserved
      reserved7 : Bool;   // Reserved
      reserved8 : Bool;   // Reserved
   END_STRUCT;
END_TYPE

TYPE "LIOLink_3SU1_IDKeySwitch_typeKeyState"
TITLE = LIOLink_3SU1_IDKeySwitch_typeKeyState
VERSION : 0.1
// Data record (index) 79 - add individually codable ID key
   STRUCT
      idByte0 : Byte;   // Byte 0 of Identification number of the individually codeable ID key
      idByte1 : Byte;   // Byte 1 of Identification number of the individually codeable ID key
      idByte2 : Byte;   // Byte 2 of Identification number of the individually codeable ID key
      idByte3 : Byte;   // Byte 3 of Identification number of the individually codeable ID key
      idByte4 : Byte;   // Byte 4 of Identification number of the individually codeable ID key
      authorizationLevel : Byte;   // Authorization level
   END_STRUCT;
END_TYPE

// folder: LIOLink/Common/Device-specific data types/SIRIUS/Common

TYPE "LIOLink_typeParameterPage0"
VERSION : 0.1
   STRUCT
      masterCommand : Byte := 16#00;   // Switch the IO-Link operation mode (Fallback, Operate, Preoperate) / Umschalten des Betriebsmodus
      masterCycleTime : Byte := 16#00;   // Master Cycle Time / Zykluszeit des IO-Link Masters
      minCycleTime : Byte := 16#00;   // Minimum Device Cycle Time / Minimale Zykluszeit eines Geraetes
      frameCapability : Byte := 16#00;   // Supported frame types for communication / Unterstuetzter Typ für die Kommunikation
      ioLinkRevisionID : Byte := 16#00;   // IO-Link protocol version implemented on the device / IO-Link Protokollversion
      processDataIn : Byte := 16#00;   // Number and structure of the data process image of the inputs to the master / Prozessdatenabbild der Eingaenge
      processDataOut : Byte := 16#00;   // Number and structure of the data process image of the outputs to the master / Prozessdatenabbild der Ausgaenge
      vendorID1 : Byte := 16#00;   // Unique vendor identification number / Eindeutige Herstelleridentifikationsnummer
      vendorID2 : Byte := 16#00;   // Siemens:0x002A / Siemens = 0x002A
      deviceID1 : Byte := 16#00;   // Unique device identification number / Eindeutige Geraeteidentifikationsnummer
      deviceID2 : Byte := 16#00;   // Unique device identification number / Eindeutige Geraeteidentifikationsnummer
      deviceID3 : Byte := 16#00;   // Unique device identification number / Eindeutige Geraeteidentifikationsnummer
      functionID1 : Byte := 16#00;   // Unique function identification number / Eindeutige Funktionsidentifikationsnummer
      functionID2 : Byte := 16#00;   // Unique function identification number / Eindeutige Funktionsidentifikationsnummer
      reserved1 : Byte := 16#00;   // Reserved / Reserviert
      reserved2 : Byte := 16#00;   // Reserved / Reserviert
   END_STRUCT;
END_TYPE

// folder: LIOLink/Common/Device-specific data types/SIRIUS/SIRIUS 3UG48/3UG481x

TYPE "LIOLink_3UG481_typeMeasure"
TITLE = LIOLink_3UG481_typeMeasure
VERSION : 0.1
// Data set (index) 94 (measured values)
   STRUCT
      reserved : Array[0..15] of Byte;   // Reserved
      voltageL1L2 : Word;   // (only 3UG4815) Voltage U L1-L2 Min:160V Max:690V
      voltageL2L3 : Word;   // (only 3UG4815) Voltage U L2-L3 Min:160V Max:690V
      voltageLxL1 : Word;   // (only 3UG4815) Voltage U L3-L1 Min:160V Max:690V
      voltageLxLyMin : Word;   // (only 3UG4815) Voltage U Lx-Ly min Min:160V Max:690V
      voltageLxLyMax : Word;   // (only 3UG4815) Voltage U Lx-Ly max Min:160V Max:690V
      voltageL1N : Word;   // (only 3UG4816) Voltage U L1-N Min:90V Max:400V
      voltageL2N : Word;   // (only 3UG4816) Voltage U L2-N Min:90V Max:400V
      voltageL3N : Word;   // (only 3UG4816) Voltage U L3-N Min:90V Max:400V
      voltageLxNmin : Word;   // (only 3UG4816) Voltage U Lx-N min Min:90V Max:400V
      voltageLxNmax : Word;   // (only 3UG4816) Voltage U Lx-N max Min:90V Max:400V
      asymmetry : Word;   // Asymmetry Min:0% Max:20%
   END_STRUCT;
END_TYPE

TYPE "LIOLink_3UG481_typeParam"
TITLE = LIOLink_3UG481_typeParam
VERSION : 0.1
// Data set (index) 131 (parameters)
   STRUCT
      reserved : Array[0..15] of Byte;   // Reserved
      groupDiagnostics : Bool := TRUE;   // Group diagnostics: Default: true, false; disabled, true: enabled
      groupErrorDiagnostics : Bool := TRUE;   // Group error diagnostics: Default: true, false; disabled, true: enabled
      reserved1 : Bool;   // Reserved
      reserved2 : Bool;   // Reserved
      localLimitChange : Bool := TRUE;   // Local threshold change: Default: true, false; disabled, true: enabled
      localParameterChange : Bool := TRUE;   // Local parameter change: Default: true, false; disabled, true: enabled
      localReset : Bool := TRUE;   // Local reset: Default: true, false; disabled, true: enabled
      retentiveErrorMemory : Bool;   // Retentive error memory: Default: false, false; disabled, true: enabled
      analogValueCoding : Byte := 16#30;   // Analog value coding: Default: 48, Min: 0(disabled), Max: 255
      reserved3 : Array[18..23] of Byte;   // Reserved
      resetResponse : Byte := 16#01;   // Reset response: Default: 16#01, 16#00: manual, 16#01: automatic
      delayOn : Bool := TRUE;   // Stabilzation delay (at Power ON): Default: true, false: disabled, true: enabled
      delayOn0 : Bool;   // False
      delayReset : Bool := TRUE;   // Stabilzation delay (at manual reset): Default: true, false: disabled, true: enabled
      delayReset0 : Bool;   // False
      reserved4 : Bool;   // Reserved
      reserved5 : Bool;   // Reserved
      reserved6 : Bool;   // Reserved
      reserved7 : Bool;   // Reserved
      phaseSequence : Byte := 16#04;   // Phase sequence monitoring: Default: 16#04, 16#00: disabled, 16#04: enabled - Bit 2 in Byte
      reserved14 : Byte;   // Reserved
      delayTimeStabilization : Int;   // Stabilization delay: Resolution: 0.1s=1, Default: 0, Min: 0.1s or 0s (disabled), Max: 999.9s
      delayTimeTripUp : Int;   // Stabilization delay(voltg ovrshoot): Resolution: 0.1s=1, Default: 0s, Min: 0.1s or 0s, Max: 999.9s
      delayTimeTripDown : Int;   // Stabilization delay(voltg undrshoot): Resolution: 0.1s=1, Default: 0s, Min: 0.1s or 0s, Max: 999.9s
      delayTimeTripAsymmetry : Int;   // Stabilization delay(asymmetry): Resolution: 0.1s=1, Default: 0s, Min: 0.1s or 0s, Max: 999.9s
      tresholdUp : Int;   // Threshold for overshoot: Resolution: 0.1V=1, Default:425/245V,Min: 160/90V or 0V, Max: 690/400V
      tresholdDown : Int;   // Threshold for undershoot: Resolution: 0.1V=1, Default: 375/215V, Min: 160/90V or 0V ,Max: 690/400V
      tresholdAsymmetry : Int := 50;   // Threshold for asymmetry: Resolution: 0.1%=1, Default: 5%, Min: 0.1% or 0% , Max: 20%
      warningTresholdUp : Int;   // Warng threshold for overshoot: Resolution: 0.1V=1, Default: 425/245V, Min: 160/90V or .0V, Max: 690/400V
      warningTresholdDown : Int;   // Warng threshold for undershoot:Resolution: 0.1V=1, Default: 375/215V, Min: 160/90V or0V ,Max: 690/400V
      warningTresholdAsymmetry : Int := 50;   // Warning threshold for asymmetry: Resolution: 0.1%=1, Default: 5%, Min: 0.1% or 0% , Max: 20%
      reserved15 : Array[48..53] of Byte;   // Reserved
      hysteresis : Int;   // Hysteresis: Resolution: 0.1V=1, Default: 5V, Min: 0.1V or 0V (disabled), Max: 20V
      hysteresisAsymmetry : Int;   // Hysteresis (asymmetry): Resolution: 0.1%=1, Default: 2%, Min: 0.1% or 0%, Max=5%
      responseRelay : Byte;   // Relay switching response:Default: 16#00, 16#00: Closed-circuit (NC), 16#01: Open-circuit(NO)
      reserved16 : Byte;   // Reserved
   END_STRUCT;
END_TYPE

TYPE "LIOLink_3UG481_typeDiag"
TITLE = LIOLink_3UG481_typeDiag
VERSION : 0.1
// Data set (index) 92 - diagnostics
   STRUCT
      reserved : Array[0..15] of Byte;   // Reserved
      ready : Bool;   // Read
      groupError : Bool;   // Group error
      groupWarning : Bool;   // Group warning
      reserved1 : Bool;   // Reserved
      reserved2 : Bool;   // Reserved
      parameterAssign : Bool;   // Parameter assignment active
      parameterInvalid : Bool;   // Invalid parameter
      internalError : Bool;   // Self-test error/internal error
      reserved3 : Byte;   // Reserved
      errorNumber : Word;   // Parameter error number
      reserved4 : Array[20..25] of Byte;   // Reserved
      delayTimeRunning : Bool;   // Stabilization delay running
      delayLevelUp : Bool;   // Tripping delay time running (threshold for overshoot)
      delayLevelDown : Bool;   // Tripping delay time running (threshold for undershoot)
      delayAsymmetry : Bool;   // Tripping delay time running (threshold for voltage asymmetry)
      reserved5 : Bool;   // Reserved
      reserved6 : Bool;   // Reserved
      reserved7 : Bool;   // Reserved
      reserved8 : Bool;   // Reserved
      levelUp : Bool;   // Threshold for overshoot exceeded
      levelDown : Bool;   // Threshold for undershoot violated
      voltageAsymmetry : Bool;   // Threshold for voltage asymmetry exceeded
      warningLevelUp : Bool;   // Warning threshold for overshoot exceeded
      warningLevelDown : Bool;   // Warning threshold for undershoot violated
      warningVoltageAsymmetry : Bool;   // Warning threshold for voltage asymmetry exceeded
      reserved9 : Bool;   // Reserved
      reserved10 : Bool;   // Reserved
      reserved11 : Bool;   // Reserved
      phaseFailureL1 : Bool;   // Phase failure L1
      phaseFailureL2 : Bool;   // Phase failure L2
      phaseFailureL3 : Bool;   // Phase failure L3
      phaseFailureN : Bool;   // Phase failure N conductor
      phaseSeqL1L2L3 : Bool;   // Phase sequence L1-L2-L3
      phaseSeqL3L2L1 : Bool;   // Phase sequence L3-L2-L1
      phaseSeqError : Bool;   // Phase sequence error
      reserved12 : Byte;   // Reserved
   END_STRUCT;
END_TYPE

TYPE "LIOLink_3UG481_typeAll"
TITLE = LIOLink_3UG481_typeAll
VERSION : 0.1
// Contains all the information about 3UG481
   STRUCT
      parameterPage0 : "LIOLink_typeParameterPage0";   // ID0: Parameter page 0
      systemCommands : Byte;   // ID2: System Commands (0x80 for device reset, 0x82 for factory reset)
      vendorName : String[11];   // ID16: Vendor name
      vendorText : String[64];   // ID17: Vendor text
      productName : String[64];   // ID18: Product name
      productID : String[14];   // ID19: Product ID
      hwRevision : String[7];   // ID22: Hardware revision
      fwRevision : String[7];   // ID23: Firmware revision
      appSpecificName : String[32];   // ID24: Application specific name
      diagnostics : "LIOLink_3UG481_typeDiag";   // ID92: Diagnostics
      measuredValues : "LIOLink_3UG481_typeMeasure";   // ID94: Measurement values
      parameters : "LIOLink_3UG481_typeParam";   // ID131: Parameters
   END_STRUCT;
END_TYPE

// folder: LIOLink/Common/Device-specific data types/SIRIUS/SIRIUS 3UG48/3UG4822

TYPE "LIOLink_3UG4822_typeMeasure"
TITLE = LIOLink_3UG4822_typeMeasure
VERSION : 0.1
// Data set (index) 94 (measured values)
   STRUCT
      reserved : Array[0..15] of Byte;   // Reserved
      currentI1Pa : Word;   // Current I1 (PA) Min:0,05A Max:10A (if trnsfrmr trnsmissn factor is deactivated)
      reserved1 : Array[18..27] of Byte;   // Reserved
      currentI1 : DWord;   // Current I1 Min:0,05A Max:10A (when transformr transmissn factor is deactivated)
      reserved2 : Array[32..51] of Byte;   // Reserved
   END_STRUCT;
END_TYPE

TYPE "LIOLink_3UG4822_typeParam"
TITLE = LIOLink_3UG4822_typeParam
VERSION : 0.1
// Data set (index) 131 (parameters)
   STRUCT
      reserved : Array[0..15] of Byte;   // Reserved
      groupDiagnostics : Bool := TRUE;   // Group diagnostics: Default: true, false; disabled, true: enabled
      groupErrorDiagnostics : Bool := TRUE;   // Group error diagnostics: Default: true, false; disabled, true: enabled
      reserved1 : Bool;   // Reserved
      reserved2 : Bool;   // Reserved
      localLimitChange : Bool := TRUE;   // Local threshold change: Default: true, false; disabled, true: enabled
      localParameterChange : Bool := TRUE;   // Local parameter change: Default: true, false; disabled, true: enabled
      localReset : Bool := TRUE;   // Local reset: Default: true, false; disabled, true: enabled
      retentiveErrorMemory : Bool;   // Retentive error memory: Default: false, false; disabled, true: enabled
      analogValueCoding : Byte := 16#10;   // Analog value coding: Default: 16, Min: 0(disabled), Max: 255
      reserved3 : Array[18..23] of Byte;   // Reserved
      resetResponse : Byte := 16#01;   // Reset response: Default: 16#01, 16#00: manual, 16#01: automatic
      delayOn : Bool := TRUE;   // ON-delay time (at Power ON): Default: true, false: disabled, true: enabled
      delayOn0 : Bool;   // False
      delayReset : Bool := TRUE;   // ON-delay time (at manual reset): Default: true, false: disabled, true: enabled
      delayReset0 : Bool;   // False
      delayRestart : Bool;   // ON-delay time (at restart): Default: true, false: disabled, true: enabled
      delayRestart0 : Bool;   // False
      reserved4 : Bool;   // Reserved
      reserved5 : Bool;   // Reserved
      delayTime : Int := 0;   // ON-delay time: Resolution: 0.1=1s, Default: 0s, Min: 0.1s or 0s (disabled), Max: 999.9s
      delayTimeTripUp : Int;   // Tripping delay time (in the case of current overshoot): Resolution: 0.1s=1, Default: 0, Min: 0.1s or 0s, Max: 999.9s
      delayTimeTripDown : Int;   // Tripping delay time (in the case of current undershoot): Resolution: 0.1s=1, Default: 0, Min: 0.1s or 0s, Max: 999.9s
      tresholdUp : DInt := 250;   // Threshold for overshoot: Resolution: 0.01A=1, Default: 2.5A, Min: 0.05A or 0A (disabled), Max: 10A
      tresholdDown : DInt := 150;   // Threshold for undershoot: Resolution: 0.01A=1, Default: 1.5A, Min: 0.05A or 0A (disabled), Max: 10A
      warningTresholdUp : DInt := 250;   // Warning threshold for overshoot: Resolution: 0.01A=1, Default: 2.5A, Min: 0.05A or 0A (disabled), Max: 10A
      warningTresholdDown : DInt := 150;   // Warning threshold for undershoot: Resolution: 0.01A=1, Default: 1.5A, Min: 0.05A or 0A (disabled), Max: 10A
      reserved7 : Array[48..55] of Byte;   // Reserved
      hysteresis : DInt := 50;   // Hysteresis: Resolution: Resolution: 0.01A=1, Default: 0,05A, Min: 0.01A or 0A (disabled), Max: 5A
      factorTransformer : Int;   // Transformer transmission factor: , Default: 0, Min: 0 or 2, Max: 750
      responseRelay : Byte;   // Relay switching response:Default: 16#00, 16#00: Closed-circuit principle NC, I > 50 mA, 16#01: Open-circuit principle NO, I > 50 mA, 16#10: Closed-circuit principle NC, Us = on, 16#11: Open-circuit principle NO, Us = on
      reserved8 : Byte;   // Reserved
   END_STRUCT;
END_TYPE

TYPE "LIOLink_3UG4822_typeDiag"
TITLE = LIOLink_3UG4822_typeDiag
VERSION : 0.1
// Data set (index) 92 - diagnostics
   STRUCT
      reserved : Array[0..15] of Byte;   // Reserved
      ready : Bool;   // Ready
      groupError : Bool;   // Group error
      groupWarning : Bool;   // Group warning
      reserved1 : Bool;   // Reserved
      reserved2 : Bool;   // Reserved
      parameterAssign : Bool;   // Parameter assignment active
      parameterInvalid : Bool;   // Invalid parameter
      internalError : Bool;   // Self-test error/internal error
      reserved3 : Byte;   // Reserved
      errorNumber : Word;   // Parameter eroor number
      reserved4 : Array[20..25] of Byte;   // Reserve
      delayTimeRunning : Bool;   // ON-delay time running
      delayLevelUp : Bool;   // Tripping delay time running (threshold for overshoot)
      delayLevelDown : Bool;   // Tripping delay time running (threshold for undershoot)
      reserved5 : Bool;   // Reserved
      reserved6 : Bool;   // Reserved
      reserved7 : Bool;   // Reserved
      reserved8 : Bool;   // Reserved
      reserved9 : Bool;   // Reserved
      levelUp : Bool;   // Threshold for overshoot exceeded
      levelDown : Bool;   // Threshold for undershoot violated
      warningLevelUp : Bool;   // Warning threshold for overshoot exceeded
      warningLevelDown : Bool;   // Warning threshold for undershoot violated
      reserved10 : Bool;   // Reserved
      reserved11 : Bool;   // Reserved
      reserved12 : Bool;   // Reserved
      reserved13 : Bool;   // Reserved
   END_STRUCT;
END_TYPE

TYPE "LIOLink_3UG4822_typeAll"
TITLE = LIOLink_3UG4822_typeAll
VERSION : 0.1
// Contains all the information about 3UG4822
   STRUCT
      parameterPage0 : "LIOLink_typeParameterPage0";   // ID0: Parameter page 0
      systemCommands : Byte;   // ID2: System Commands (0x80 for device reset, 0x82 for factory reset)
      vendorName : String[11];   // ID16: Vendor name
      vendorText : String[64];   // ID17: Vendor text
      productName : String[64];   // ID18: Product name
      productID : String[14];   // ID19: Product ID
      hwRevision : String[7];   // ID22: Hardware revision
      fwRevision : String[7];   // ID23: Firmware revision
      appSpecificName : String[32];   // ID24: Application specific name
      diagnostics : "LIOLink_3UG4822_typeDiag";   // ID92: Diagnostics
      measuredValues : "LIOLink_3UG4822_typeMeasure";   // ID94: Measurement values
      parameters : "LIOLink_3UG4822_typeParam";   // ID131: Parameters
   END_STRUCT;
END_TYPE

// folder: LIOLink/Common/Device-specific data types/SIRIUS/SIRIUS 3UG48/3UG4825

TYPE "LIOLink_3UG4825_typeMeasure"
TITLE = LIOLink_3UG4825_typeMeasure
VERSION : 0.1
// Data set (index) 94 (measured values)
   STRUCT
      reserved : Array[0..15] of Byte;   // Reserved
      residualCurrentIrPa : Word;   // Residual current Ir (PA), Min: 0,0 A, Max: 43,0 A
      residualCurrentIr : DWord;   // Residual current Ir, Min: 0,0 A, Max: 43,0 A
   END_STRUCT;
END_TYPE

